(* IEC 61131-3 sources: CS_4_Aufzugsteuerung/src/Stations/CP112/Steuerung/Class/DiasMasterMain (part 2) *)

	l.eax		  RTCY
	and.eax		Dmrealtime
	call		  StoreNewPointers

END_FUNCTION
#endif

#ifdef _LSL_TARGETARCH_ARM
FUNCTION VIRTUAL GLOBAL DiasMasterMain::AddRet
  VAR_INPUT
    RTCY		: DINT;
  END_VAR

  if (RTCY AND DMREALTIME) = DMREALTIME then
    ud_DelayRealtime += C_TimeRet;
  else
    ud_DelayCyclic += C_TimeRet;
  end_if;

  (PtrCode + IPSub + RetStruct.Opc)^ := DbRet;

  IPSub += sizeof(RetStruct);

END_FUNCTION

#else
FUNCTION AWL VIRTUAL GLOBAL DiasMasterMain::AddRet
  VAR_INPUT
    RTCY		: DINT;
  END_VAR

	l.eax		  RTCY
	and.eax		Dmrealtime

//#SR001 Start
	CMP.EAX		Dmrealtime
	JNE			  LABEL_AR_NORT
	ADD.D		  ud_DelayRealtime,C_TimeRet
  JMP       LABEL_AR_TIMETAKEN

LABEL_AR_NORT
//#SR001 End
	ADD.D		  ud_DelayCyclic,C_TimeRet

LABEL_AR_TIMETAKEN

	call		  GetProgPointer

  l.ebx     PtrCode

	l.b			  (edx+ebx+RetStruct.Opc),DbRet			     // opcode Ret
	add.edx		sizeof (RetStruct)

	l.eax		  RTCY
	and.eax		Dmrealtime
	call		  StoreNewPointers

END_FUNCTION
#endif

//[English]
// Does a 16 Bit read access
//[Globals]		_RTOSVersion			: OS version
//				_lsl_pos				: OS interface structure
//[Members]
//[Locals]		ui_data			:R/W	:intermediate storeage of data
//				di_ret			:R/W	:returnvalue of OS
//[>Adress]		Module address and offset
//[<Data]		Data read
FUNCTION VIRTUAL GLOBAL DiasMasterMain::Rd16Bit
  VAR_INPUT
    Adress	: UDINT;
  END_VAR
  VAR_OUTPUT
    Data		: DINT;
  END_VAR
  VAR
    ui_data : uint;
    di_ret	: dint;
  END_VAR

	//ws005
	//*****************************************************
	//***** use OS functions instead of own functions *****
	//*****************************************************
	if( _RTOSVersion >= OSVersionDIASIO )then
		if( p_SemaHandle <> NIL )then			//ws007
			To_Multitask.Wait( p_SemaHandle );	//ws006
		end_if;
		di_ret := OS_DIAS_ReadWord( pDIAS  := pDIAS,
								   us_mod  := ( ( Adress shr 8 ) and 16#ff )$usint,
								   ui_off  := ( Adress and 16#ff )$uint,
								   ui_data := #ui_data );
		if( p_SemaHandle <> NIL )then				//ws007
			To_Multitask.Signal( p_SemaHandle );	//ws006
		end_if;
		if( di_ret <> 0 )then
			Data := 0;
			TraceAsyncError(( ( Adress shr 8 ) and 16#ff )$usint);
		else
			Data := ui_data;
		end_if;
	else
	//*****************************************************
	//*** use own functions (should be obsolete by now) ***
	//*****************************************************
	// /ws005
		TraceAsyncError(( ( Adress shr 8 ) and 16#ff )$usint);
	end_if;

END_FUNCTION

#ifdef _LSL_TARGETARCH_ARM
FUNCTION VIRTUAL GLOBAL DiasMasterMain::AddRd32Bit
  VAR_INPUT
    Adress		  : HINT;
    RTCY		    : DINT;
    thisp		    : ^void;
    callOptions : USINT;
  END_VAR
  VAR_OUTPUT
    Handle		  : DINT;
  END_VAR

  if (RTCY AND Dmrealtime) = Dmrealtime then
    ud_DelayRealtime += C_TimeRd8Bit + 3*(C_TimeRd16Bit - C_TimeRd8Bit); // appraised value: 1*basetime + 4*time for 1 byte (instead of C_TimeRd32Bit)
    ui_RtDIASAccesses += 1;
  else
    ud_DelayCyclic += C_TimeRd8Bit + 3*(C_TimeRd16Bit - C_TimeRd8Bit); // appraised value: 1*basetime + 4*time for 1 byte (instead of C_TimeRd32Bit)
    ui_CyDIASAccesses += 1;
  end_if;

  (PtrCode + IPSub + Rd32Struct.Opc)^         := DbRd32;
  (PtrCode$^HINT + IPSub + Rd32Struct.ChAdr)^ := Adress;

  ARM_EAX := RTCY$UDINT;
  ARM_EDI := thisp$UDINT;
  GetHandle(Rd32Struct.Data, callOptions);
  Handle := ARM_EAX$DINT;
  IPSub += sizeof(Rd32Struct);

END_FUNCTION

#else
// ***************************************
//   put programm into the buffer
// ***************************************
//  this is a 16 bit read
//  the thispointer we need to call the update method
//

FUNCTION AWL VIRTUAL GLOBAL DiasMasterMain::AddRd32Bit
	VAR_INPUT
		Adress 	    : HINT;
		RTCY 	      : DINT;
		thisp 	    : ^void;
		callOptions : USINT;
	END_VAR
	VAR_OUTPUT
		Handle 	    : DINT;
	END_VAR

	l.eax		  RTCY
	and.eax		Dmrealtime

//#SR001 Start
	CMP.EAX		Dmrealtime
	JNE			  LABEL_AR32B_NORT
	ADD.D		  ud_DelayRealtime,C_TimeRd32Bit
	inc.w		  ui_RtDIASAccesses
  JMP       LABEL_AR32B_TIMETAKEN

LABEL_AR32B_NORT
	ADD.D		  ud_DelayCyclic,C_TimeRd32Bit
	inc.w		  ui_CyDIASAccesses
//#SR001 End

LABEL_AR32B_TIMETAKEN

	call		  GetProgPointer

  l.ebx     PtrCode

	l.b			  (edx+ebx+Rd32Struct.Opc),DbRd32	   			// opcode Read 8
	l.ax		  Adress					// adress lo+high
	s.ax		  (edx+ebx+Rd32Struct.ChAdr+0)

	l.ax		  RTCY+0
	l.edi		  thisp				    // to put into then handle

  push.b    callOptions

	push.d		Rd16Struct.Data			// direct pointer on the data
	call		  GetHandle

  add.esp 5

	s.eax		  Handle

	add.edx		sizeof (Rd32Struct)

	l.eax		  RTCY
	and.eax		Dmrealtime
	call		  StoreNewPointers

END_FUNCTION
#endif

#ifdef _LSL_TARGETARCH_ARM
FUNCTION VIRTUAL GLOBAL DiasMasterMain::AddRd8Bit
  VAR_INPUT
    Adress		  : HINT;
    RTCY		    : DINT;
    thisp		    : ^void;
    callOptions : USINT;
  END_VAR
  VAR_OUTPUT
    Handle		  : DINT;
  END_VAR

  if (RTCY AND Dmrealtime) = Dmrealtime then
    ud_DelayRealtime += C_TimeRd8Bit;
    ui_RtDIASAccesses += 1;
  else
    ud_DelayCyclic += C_TimeRd8Bit;
    ui_CyDIASAccesses += 1;
  end_if;

  (PtrCode + IPSub + Rd8Struct.Opc)^         := DbRd8;
  (PtrCode$^HINT + IPSub + Rd8Struct.ChAdr)^ := Adress;

  ARM_EAX := RTCY$UDINT;
  ARM_EDI := thisp$UDINT;
  GetHandle(Rd8Struct.Data, callOptions);
  Handle := ARM_EAX$DINT;
  IPSub += sizeof(Rd8Struct);

END_FUNCTION

#else
// ***************************************
//   put programm into the buffer
// ***************************************
//  this is a 8 bit read
//  the thispointer we need to call the update method
//

FUNCTION AWL VIRTUAL GLOBAL DiasMasterMain::AddRd8Bit
	VAR_INPUT
		Adress 	    : HINT;
		RTCY 	      : DINT;
		thisp 	    : ^void;
		callOptions : USINT;
	END_VAR
	VAR_OUTPUT
		Handle 	    : DINT;
	END_VAR

	l.eax		  RTCY
	and.eax		Dmrealtime

//#SR001 Start
	CMP.EAX		Dmrealtime
	JNE			  LABEL_AR8B_NORT
	ADD.D		  ud_DelayRealtime,C_TimeRd8Bit
	inc.w		  ui_RtDIASAccesses			//#SR021
  JMP       LABEL_AR8B_TIMETAKEN

LABEL_AR8B_NORT
	ADD.D		  ud_DelayCyclic,C_TimeRd8Bit
	inc.w		  ui_CyDIASAccesses
//#SR001 End

LABEL_AR8B_TIMETAKEN

	call		  GetProgPointer

  l.ebx     PtrCode

	l.b			  (edx+ebx+Rd8Struct.Opc),DbRd8	   			// opcode Read 8
	l.ax		  Adress					// adress lo+high
	s.ax		  (edx+ebx+Rd8Struct.ChAdr+0)

	l.ax		  RTCY+0
	l.edi		  thisp				    // to put into then handle

  push.b    callOptions

	push.d		Rd8Struct.Data			// direct pointer on the data
	call		  GetHandle

  add.esp   5

	s.eax		  Handle
	add.edx		sizeof (Rd8Struct)

	l.eax		  RTCY
	and.eax		Dmrealtime
	call		  StoreNewPointers

END_FUNCTION
#endif

#ifdef _LSL_TARGETARCH_ARM
FUNCTION VIRTUAL GLOBAL DiasMasterMain::AddRTBSync
  VAR_INPUT
    Adress		: HINT;
  END_VAR
  VAR_OUTPUT
    FirstRTB	: DINT;
  END_VAR
  #ifdef OldDiasXilinx
  VAR
    pUSINT : ^USINT;
  END_VAR
#endif

  FirstRTB := 0;

  if DiasType <> 2 then

#IFNDEF OldDiasXilinx
    if RTBSyncAdr = NIL then
      RTBSyncAdr := (16#100*63+16#8002)$^USINT;// global sync

      FirstRTB := 1;
    end_if;
#ELSE
    if NumberSyncs >= NumberLocalSyncs then
      ErrorLocalSyncTrace();
    else
      ((#RtbLocalSyncAdr)$^DINT + NumberSyncs * (SIZEOF(RtbLocalSyncAdr)/NumberLocalSyncs))^ := Adress + 16#8000;
    end_if;
#ENDIF
  else
    // DiasType = 2 --> it is a new Master
#IFNDEF OldDiasXilinx
    if (SyncProgPtr + CntrlStruct.OPC)^ <> DbCntrl then
      (SyncProgPtr + CntrlStruct.OPC)^          := DbCntrl;
      (SyncProgPtr$^UINT + CntrlStruct.chAdr)^  := 16#100*63+2;
      (SyncProgPtr + CntrlStruct.Data)^         := 0;
      FirstRTB := 1;

      ud_DelayRealtime := ud_DelayRealtime + C_TimeControlWrite - C_TimeNop * 4; //because the 4 Nops were overwritten
    end_if;
#ELSE
    if NumberSyncs >= NumberLocalSyncs then
      ErrorLocalSyncTrace();
    else
      pUSINT := #CallsRt[0] + sizeof(TmrStruct) + NumberSyncs * SIZEOF(CntrlStruct);

      if (pUSINT + CntrlStruct.OPC)^ <> DbCntrl then
        (pUSINT + CntrlStruct.OPC)^         := DbCntrl;
        (pUSINT$^UINT + CntrlStruct.chAdr)^ := Adress;
        (pUSINT + CntrlStruct.Data)^        := 0;

        ud_DelayRealtime := ud_DelayRealtime + C_TimeControlWrite - C_TimeNop * 4; //because the 4 Nops were overwritten
      end_if;
    end_if;
#ENDIF
  end_if;

  NumberSyncs += 1;

  if FirstRTB = 1 then
    us_SyncModule := (Adress SHR 8)$USINT;
  end_if;

END_FUNCTION

#else

// *************************************************
//   RTB is fixed reserved for one MODUL
// *************************************************
//
//  if FirstRTB <> 0 then this modul is the first with RTB
//  and has to do perhaps something special
//  if FirstRTB = 0 then it already exists a modul with RTBSYNC
//

FUNCTION AWL VIRTUAL GLOBAL DiasMasterMain::AddRTBSync
  VAR_INPUT
    Adress		: HINT;
  END_VAR
  VAR_OUTPUT
    FirstRTB	: DINT;
  END_VAR

	l.d			FirstRTB,0

	cmp.b		DiasType,2			//ws005
	je			AddRTBIMaster		// --> it is a new Master

#IFNDEF OldDiasXilinx
	cmp.d		RTBSyncAdr,0
	jne			AddRTBSyncRet

	L.EDI		16#100*63+16#8002 		// global sync  //ws005: faster

	s.edi		RTBSyncAdr

	l.d			FirstRTB,1						// first RTB
#ELSE
	LZXW.EDI	Adress
	ADD.EDI		16#8000

	LZXB.EAX	NumberSyncs
	CMP.AL		NumberLocalSyncs
	JAE			  ErrorSync
	L.AH		  SIZEOF(RtbLocalSyncAdr)/NumberLocalSyncs
	MUL			  AH
	ADD.EAX		#RtbLocalSyncAdr

	S.EDI		  (EAX)
#ENDIF
	jmp			  AddRTBSyncRet

AddRTBIMaster
#IFNDEF OldDiasXilinx

	//#SR003 Start
	l.edi	    SyncProgPtr
	//#SR003 End

	cmp.b		  (edi+CntrlStruct.OPC),DbCntrl
	je			  AddRTBSyncRet

	l.b			  (edi+CntrlStruct.OPC),DbCntrl

	l.ax		  16#100*63+2 		// global sync

	s.ax		  (edi+CntrlStruct.chAdr+0)		// the modul normal = 63 (global SYNC)

	l.b			  (edi+CntrlStruct.Data),0		// we always write data 0
	l.d			  FirstRTB,1						// first RTB

//#SR001 Start
	SUB.D		  ud_DelayRealtime,C_TimeNop * 4			//because the 4 Nops were write over
	ADD.D		  ud_DelayRealtime,C_TimeControlWrite
//#SR001 End

#ELSE
	l.edi		  #CallsRt
	add.edi		sizeof (TmrStruct)  // the first INSTR is tmr

	LZXB.EAX	NumberSyncs
	CMP.AL		NumberLocalSyncs
	JAE			  ErrorSync
	L.AH		  SIZEOF(CntrlStruct)
	MUL			  AH
	ADD.EDI		EAX

	cmp.b		  (edi+CntrlStruct.OPC),DbCntrl
	je			  AddRTBSyncRet

	l.b			  (edi+CntrlStruct.OPC),DbCntrl
	l.ax		  Adress
	s.ax		  (edi+CntrlStruct.chAdr+0)		// the modul normal = 63 (global SYNC)

	l.b			  (edi+CntrlStruct.Data),0		// we always write data 0

//#SR001 Start
	SUB.D		  ud_DelayRealtime,C_TimeNop * 4			//because the 4 Nops were write over
	ADD.D		  ud_DelayRealtime,C_TimeControlWrite
//#SR001 End

	JMP			  AddRTBSyncRet

ErrorSync
	FC			  ErrorLocalSyncTrace
#ENDIF

AddRTBSyncRet

	INC.B		  NumberSyncs

	//#SR008 start
	cmp.d		  FirstRTB,1
	jne			  LABEL_End

	l.ax		  Adress
	shr.ax		8
	s.al		  us_SyncModule

LABEL_End
	//#SR008 end

END_FUNCTION
#endif

#ifdef _LSL_TARGETARCH_ARM
FUNCTION VIRTUAL GLOBAL DiasMasterMain::AddWR16Bit
  VAR_INPUT
    adress	    : Hint;
    RTCY		    : DINT;
    thisp		    : ^void;
    data		    : UINT;
    callOptions : USINT;
  END_VAR
  VAR_OUTPUT
    handle		  : DINT;
  END_VAR

  if (RTCY AND Dmrealtime) = Dmrealtime then
    ud_DelayRealtime += C_TimeWr16Bit;
    ui_RtDIASAccesses += 1;
  else
    ud_DelayCyclic += C_TimeWr16Bit;
    ui_CyDIASAccesses += 1;
  end_if;

  (PtrCode + IPSub + Wr16Struct.Opc)^         := DbWr16;
  (PtrCode$^HINT + IPSub + Wr16Struct.ChAdr)^ := Adress;
  (PtrCode$^HINT + IPSub + Wr16Struct.Data)^  := data;

  ARM_EAX := RTCY$UDINT;
  ARM_EDI := thisp$UDINT;
  GetHandle(Wr16Struct.Data, callOptions);
  Handle := ARM_EAX$DINT;
  IPSub += sizeof(Wr16Struct);

END_FUNCTION

// ***************************************
//   put programm into the buffer
// ***************************************
//  this is a 16 bit read
//  the thispointer we need to call the update method
//
#else
FUNCTION AWL VIRTUAL GLOBAL DiasMasterMain::AddWR16Bit
	VAR_INPUT
		adress 	      : HINT;
		RTCY 	        : DINT;
		thisp 	      : ^void;
		data 	        : UINT;
		callOptions 	: USINT;
	END_VAR
	VAR_OUTPUT
		handle 	      : DINT;
	END_VAR

	l.eax		  RTCY
	and.eax		Dmrealtime

//#SR001 Start
	CMP.EAX		Dmrealtime
	JNE			  LABEL_AW16B_NORT
	ADD.D		  ud_DelayRealtime,C_TimeWr16Bit
	inc.w		  ui_RtDIASAccesses			//#SR021
  JMP       LABEL_AW16B_TIMETAKEN

LABEL_AW16B_NORT
	ADD.D		  ud_DelayCyclic,C_TimeWr16Bit
	inc.w		  ui_CyDIASAccesses
//#SR001 End

LABEL_AW16B_TIMETAKEN

	call		  GetProgPointer

  l.ebx     PtrCode

	l.b			  (edx+ebx+Wr16Struct.Opc),DbWr16	   			// opcode Read 8
	l.ax		  Adress					// adress lo+high
	s.ax		  (edx+ebx+Wr16Struct.ChAdr+0)

	l.ax		  data
	s.ax		  (edx+ebx+Wr16Struct.Data)

	l.ax		  RTCY+0
	l.edi		  thisp				    // to put into then handle

  push.b    callOptions

	push.d		Wr16Struct.Data			// direct pointer on the data
	call		  GetHandle

  add.esp   5

	s.eax		  Handle

	add.edx		sizeof (Wr16Struct)
	l.eax		  RTCY
	and.eax		Dmrealtime
	call		  StoreNewPointers

END_FUNCTION
#endif

#ifdef _LSL_TARGETARCH_ARM
FUNCTION VIRTUAL GLOBAL DiasMasterMain::AddWr8Bit
	VAR_INPUT
		adress 	    : HINT;
		RTCY 	      : DINT;
		thisp 	    : ^void;
		Data 	      : USINT;
		callOptions : USINT;
	END_VAR
	VAR_OUTPUT
		Handle 	    : DINT;
	END_VAR

  if (RTCY AND Dmrealtime) = Dmrealtime then
    ud_DelayRealtime += C_TimeWr8Bit;
    ui_RtDIASAccesses += 1;
  else
    ud_DelayCyclic += C_TimeWr8Bit;
    ui_CyDIASAccesses += 1;
  end_if;

  (PtrCode + IPSub + Wr8Struct.Opc)^         := DbWr8;
  (PtrCode$^HINT + IPSub + Wr8Struct.ChAdr)^ := Adress;
  (PtrCode$^HINT + IPSub + Wr8Struct.Data)^  := data;

  ARM_EAX := RTCY$UDINT;
  ARM_EDI := thisp$UDINT;
  GetHandle(Wr8Struct.Data, callOptions);
  Handle := ARM_EAX$DINT;
  IPSub += sizeof(Wr8Struct);

END_FUNCTION

#else
FUNCTION AWL VIRTUAL GLOBAL DiasMasterMain::AddWr8Bit
	VAR_INPUT
		adress 	    : HINT;
		RTCY 	      : DINT;
		thisp 	    : ^void;
		Data 	      : USINT;
		callOptions : USINT;
	END_VAR
	VAR_OUTPUT
		Handle 	    : DINT;
	END_VAR

	l.eax		  RTCY
	and.eax		Dmrealtime

//#SR001 Start
	CMP.EAX		Dmrealtime
	JNE			  LABEL_AW8B_NORT
	ADD.D		  ud_DelayRealtime,C_TimeWr8Bit
	inc.w		  ui_RtDIASAccesses			//#SR021
  JMP       LABEL_AW8B_TIMETAKEN

LABEL_AW8B_NORT
	ADD.D		  ud_DelayCyclic,C_TimeWr8Bit
	inc.w		  ui_CyDIASAccesses
//#SR001 End

LABEL_AW8B_TIMETAKEN

	call		  GetProgPointer

  l.ebx     PtrCode

	l.b			  (edx+ebx+Wr8Struct.Opc),DbWr8	   			// opcode Read 8
	l.ax		  Adress					// adress lo+high
	s.ax		  (edx+ebx+Wr8Struct.ChAdr+0)
	l.al		  data
	s.al		  (edx+ebx+Wr8Struct.Data)

	l.ax		  RTCY+0
	l.edi		  thisp				    // to put into then handle

  push.b    callOptions

	push.d	  Wr8Struct.Data			// direct pointer on the data
	call		  GetHandle

  add.esp   5
	s.eax		  Handle

	add.edx		sizeof (Wr8Struct)

	l.eax		  RTCY
	and.eax		Dmrealtime
	call		  StoreNewPointers

END_FUNCTION
#endif

//[English]
// Function is writing into controlarea of a diasmodul
//[Globals]		_RTOSVersion		: OS version
//				_lsl_pos			: OS interface structure
//[Members]
//[Locals]
//[>Adress]		High Byte Modulnumber, Low Byte offset in Controlarea
//[>Data]		Data to write
//[<state]		0..success
FUNCTION VIRTUAL GLOBAL DiasMasterMain::WrCntr
  VAR_INPUT
    adress		: DINT;
    Data		  : Usint;
  END_VAR
  VAR_OUTPUT
    state		: DINT;
  END_VAR

	//ws005
	//*****************************************************
	//***** use OS functions instead of own functions *****
	//*****************************************************
	if( _RTOSVersion >= OSVersionDIASIO )then
		if( p_SemaHandle <> NIL )then			//ws007
			To_Multitask.Wait( p_SemaHandle );	//ws006
		end_if;
		state := OS_DIAS_WriteCtrl_( pDIAS  := pDIAS,
									us_mod  := ( ( Adress shr 8 ) and 16#ff )$usint,
									ui_off  := ( Adress and 16#ff )$uint,
									us_data := Data );
		if( p_SemaHandle <> NIL )then				//ws007
			To_Multitask.Signal( p_SemaHandle );	//ws006
		end_if;
		if( state <> 0 )then
			TraceAsyncError(( ( Adress shr 8 ) and 16#ff )$usint);
		end_if;
	else
	//*****************************************************
	//*** use own functions (should be obsolete by now) ***
	//*****************************************************
		if( ( _WhoAmI = 16#19 ) | ( _WhoAmI = 16#17 ) )then //ET261 and ETT321
			state := OS_DIAS_WriteCtrl_( pDIAS  := pDIAS,
										us_mod  := ( ( Adress shr 8 ) and 16#ff )$usint,
										ui_off  := ( Adress and 16#ff )$uint,
										us_data := Data );
			if( state <> 0 )then
				TraceAsyncError(( ( Adress shr 8 ) and 16#ff )$usint);
			end_if;
		else

	// /ws005
			TraceAsyncError(( ( Adress shr 8 ) and 16#ff )$usint);
		end_if;
	end_if;

END_FUNCTION
//[#ENGLISH]
//[>Time_uSec]Time in uSec (valid from 0-255)

#ifdef _LSL_TARGETARCH_ARM
FUNCTION VIRTUAL GLOBAL DiasMasterMain::AddWait
  VAR_INPUT
    RTCY		  : DINT;
    Time_uSec	: DINT;
  END_VAR

  if (RTCY AND Dmrealtime) = Dmrealtime then
    ud_DelayRealtime += Time_uSec$UDINT * 1000;
  else
    ud_DelayCyclic += Time_uSec$UDINT * 1000;
  end_if;

  (PtrCode + IPSub + DelayStruct.Opc)^       := DbDelay;
  (PtrCode + IPSub + DelayStruct.TIME_uSec)^ := Time_uSec$HSINT;

  IPSub += sizeof(DelayStruct);

END_FUNCTION
#else

FUNCTION AWL VIRTUAL GLOBAL DiasMasterMain::AddWait
  VAR_INPUT
    RTCY		  : DINT;
    Time_uSec	: DINT;
  END_VAR

	l.eax		  RTCY
	and.eax		Dmrealtime

//#SR001 Start
	l.ecx		  Time_usec
	imul.ecx	ecx,1000
	CMP.EAX		Dmrealtime
	JNE			  LABEL_AW_NORT
	ADD.D		  ud_DelayRealtime,ecx
  JMP       LABEL_AW_TIMETAKEN

LABEL_AW_NORT
  ADD.D		  ud_DelayCyclic,ecx
//#SR001 End

LABEL_AW_TIMETAKEN

	call		  GetProgPointer

  l.ebx     PtrCode

	l.b			  (edx+ebx+DelayStruct.OPC),DbDelay	   			// opcode delay uSec
	l.eax		  Time_uSec
	s.al		  (edx+ebx+DelayStruct.TIME_uSec)
	add.edx		sizeof (DelayStruct)

	l.eax		  RTCY
	and.eax		Dmrealtime
	call		  StoreNewPointers

END_FUNCTION
#endif

FUNCTION VIRTUAL GLOBAL DiasMasterMain::GetPllTime
  VAR_OUTPUT
    PllTime		: DINT;
  END_VAR
  VAR
    objinfo : LSLOBJ_INFO;
    Val		: DINT;
  END_VAR

	IF PllTimeGlob = 0 THEN

		To_TaskObjectControl.GetObjectInfo(this,OBJ_RT,#objinfo);			//#SR009

		// the set value of object
		PllTimeGlob := objinfo.period$DINT;
		IF PllTimeGlob = 0 THEN
#ifdef HWC_LogError
      HWC_LogError(this, "@0002 (DiasMasterMain::GetPllTime) A realtime of object 'DiasMasterC' is required !! ( 1ms is the default value ) !!");
#else
      TRACE("A realtime of object 'DiasMasterC' is required !! ( 1ms is the default value ) !!");
#endif
		END_IF;

    //look if we have µs or ms (µs msb is set)
    if ( ( objinfo.period and 16#8000_0000 ) = 0 ) then

      //we need our task time in µs
      ud_TaskTime := objinfo.period * 1000;
    else

      //we have already µs seconds
      ud_TaskTime := objinfo.period and 16#7FFF_FFFF;
    end_if;

		//#SR013 start
		us_RtPasses := 1;
		us_ModuleUpdate1ms := 1;
		us_MuSecMode := 0;

		//look if we have no old OS ( from 1.1.50 upwards)
		if _RtOSversion >= 16#1132 then
			//RTOS variable _ClockTicks ( with pointer because of linker error with old loaders without this variable)
			//_Firstscan has Offset 0EB8 and _ClockTicks has offset 0EAB, therefore -13
			ui_ClockTicks := ( ( #_Firstscan - 13 )$^UINT )^;

      if ui_ClockTicks < 1000 then
        //is DiasMaster rt time same as OS-Time (maintimer)
        if ( PllTimeGlob and 16#7FFF_FFFF ) = ui_ClockTicks then
          // check if maintimer has a valid value
          if ( 1000 mod ui_ClockTicks ) | ui_ClockTicks < 50 then
#ifdef HWC_LogError
            HWC_LogError(this, "@0003 (DiasMasterMain::GetPllTime) No valid maintimer value in OS (valid: 50,100,125,200,250,500,1000)! Master is set off!");
#else
            TRACE( "No valid maintimer value in OS (valid: 50,100,125,200,250,500,1000)! Master is set off!" );
#endif
            MasterOn := 0;
            ImOff := 1;
          else
            us_RtPasses := ( 1000 / ui_ClockTicks )$USINT;
            us_MuSecMode := 1;
            us_ModuleUpdate1ms := 0;
          end_if;
        else
          // there is only one FPGA SyncOut for OS-RT and DiasMaster, so they have to be at the same cycle
#ifdef HWC_LogError
          HWC_LogError(this, "@0004 (DiasMasterMain::GetPllTime) Rt-Time of DiasMasterC not the same as Base Rt-Time of OS (Maintimer). Master is set off!");
#else
          TRACE( "Rt-Time of DiasMasterC not the same as Base Rt-Time of OS (Maintimer). Master is set off!" );
#endif
          MasterOn := 0;
          ImOff := 1;
        end_if;
      end_if;
		end_if;
		//#SR013 End

		// but it could be a CPU with 3ms
		Val := PllTimeGlob MOD Ops.RtInterv_mSec$DINT;
		IF Val THEN
			PllTimeGlob += Ops.RtInterv_mSec$DINT - Val ;
		END_IF;

		// there could be a error
		IF PllTimeGlob < Ops.RtInterv_mSec$DINT THEN
			PllTimeGlob := Ops.RtInterv_mSec$DINT;
		END_IF;

#ifdef HWC_LogValue1
    HWC_LogValue1(this, "@0500 (DiasMasterMain::GetPllTime) PllTime = {0}", PllTimeGlob$UDINT);
#else
		//#SR008 start
		if p_KernelLog <> NIL then
			OS_KernelLog1( "DiasMaster: PllTime = %d", PllTimeGlob );
		end_if;
		//#SR008 end
#endif

		sd_PllTimeGlob_us := PllTimeGlob * 1000;		//#SR009
	END_IF;

	// aber eigentlich hängt er ja am TASK0 => #FA fragen !! => Ops.RtInterv_mSec

	PllTime := PllTimeGlob;

END_FUNCTION
//[English]
// Does a 8 Bit write access
//[Globals]		_RTOSVersion		: OS version
//				_lsl_pos			: OS interface structure
//[Members]
//[Locals]
//[>Adress]		Module address and offset
//[>Data]		Data to write
//[<State]
FUNCTION VIRTUAL GLOBAL DiasMasterMain::Wr8Bit
  VAR_INPUT
    Adress	: UDINT;
    Data		: Usint;
  END_VAR
  VAR_OUTPUT
    State		: DINT;
  END_VAR

	//ws005
	//*****************************************************
	//***** use OS functions instead of own functions *****
	//*****************************************************
	if( _RTOSVersion >= OSVersionDIASIO )then
		if( p_SemaHandle <> NIL )then			//ws007
			To_Multitask.Wait( p_SemaHandle );	//ws006
		end_if;
		State := OS_DIAS_WriteByte(pDIAS   := pDIAS,
                               us_mod  := ( ( Adress shr 8 ) and 16#ff )$usint,
                               ui_off  := ( Adress and 16#ff )$uint,
                               us_data := Data );
		if( p_SemaHandle <> NIL )then				//ws007
			To_Multitask.Signal( p_SemaHandle );	//ws006
		end_if;
		if( State <> 0 )then
			TraceAsyncError(( ( Adress shr 8 ) and 16#ff )$usint);
		end_if;
	else
	//*****************************************************
	//*** use own functions (should be obsolete by now) ***
	//*****************************************************
	// /ws005
		TraceAsyncError(( ( Adress shr 8 ) and 16#ff )$usint);
	end_if;

END_FUNCTION

FUNCTION  DiasMasterMain::DiasMasterMain
  VAR_OUTPUT
    ret_code		: CONFSTATES;
  END_VAR
  VAR
    MyProgPtr       : ^USINT;
    P2Cil		        : ^s_DiasInfoType;	//ws003
    i		            : USINT;
    PTRWDDIAS	      : ^USINT;
    SigmaTekDevInfo : ^PCICONFDATA;
    timex		        : UDINT;
#ifndef HWC_LogInit
    P2SSR		        : ^LSL_SSR;				//#SR008
#endif
    p_Obj           : ^Obj;
    p_ClsHdr        : ^ClsHdr;
    b_IsLocalMaster : BOOL;
  END_VAR

  // check if we are any kind of derivation that makes us no local master!
  b_IsLocalMaster := TRUE;
  p_Obj		:= LSL_GetHdr(this);
  p_ClsHdr := p_Obj^.pClsHdr;
  WHILE p_clsHdr^.pBaseCls <> NIL DO // go down until there is no base - we might be derived by the user....
    #pragma warning(disable: 137 )
    IF  _strcmp(str1:=#p_ClsHdr^.pDsc^.Name.Text$CHAR, str2:="Dias2DataMover") = 0
      | _strcmp(str1:=#p_ClsHdr^.pDsc^.Name.Text$CHAR, str2:="DiasMasterSplitter") = 0
      | _strcmp(str1:=#p_ClsHdr^.pDsc^.Name.Text$CHAR, str2:="DiasMasterC_Dummy") = 0 THEN
      //if we find a derivation during going down that is called Dias2DataMover or DiasMasterSplitter
      //this is no local DiasMaster and we do not need to initialize it
      b_IsLocalMaster := FALSE;
      EXIT;
    END_IF;
    #pragma warning(default: 137 )
    p_ClsHdr := p_ClsHdr^.pBaseCls;
  END_WHILE;

  MasterON := 1;
  RTBSyncAdr :=NIL;
  CDiasType:=0;
  DiasType := 16#ff;
  ud_DelayRealtime := 0;	//#SR001
  us_SyncModule := 255;	//#SR012

  //#SR013 start
  us_RtPasses := 1;
  us_ModuleUpdate1ms := 1;
  us_MuSecMode := 0;
  //#SR013 end

  PtrCY 	 := #CallsCY[0];
  IPMainCY := 0;   // stops with a end programm
  IPSub  := 0;//(DmCallRes* sizeof (CallStruct)) + sizeof (EndStruct);

  PtrRT 	 := #CallsRT[0];

  PtrCode  := #CodeRtCy[0];

  IF b_IsLocalMaster THEN

    pDIAS := _lsl_pos^.piDias;  //ws005: prepare the DIAS pointer (faster)

#ifdef HWC_LogInit
    HWC_LogInit();
#else
    //#SR008 start
    if OS_CILGET( "SSR", #P2SSR ) then
      p_KernelLog := NIL;
    else
      p_KernelLog := ( P2SSR^.KernelLog )$^DINT;
    end_if;
    //#SR008
#endif

    // test if interface already exist
    if OS_CILGET("DiasInfo", #P2Cil) then
      if ((_IOsegment$DINT <> 0) & (_IOsegment$DINT <> 16#D0000)) then
        release :=0;
        DiasType:=1;
      end_if;
    else
      DiasType := P2Cil^.DiasType$usint;
      _IOSegment$^USINT := DiasHwPointer  := P2Cil^.DiasHWPointer$^usint; //ws003
      CDiasHwPointer := P2Cil^.CDiasHWPointer$^usint;	//ws003
      CDiasType := ( P2Cil^.CDiasType )$USINT;	//ws003

      IF CDiasType = 1 THEN

        //--- CCL -----------------------------------------------------
        IF OS_CILGET("CDIAS_IRQ",#lsl_cdias_irq) = SYS_ERR_NONE THEN
          CDiasIRQpossible := 1;
        END_IF;

      ELSIF CDiasType = 2 THEN

        //--- CIPC ----------------------------------------------------
        IF OS_CILGET("CDIAS_IRQ",#lsl_cdias_irq) = SYS_ERR_NONE THEN
          CDiasIRQpossible := 1;
        END_IF;

        IF OS_CILGET("PCICONFIG", #pSPCIInfo) =  SYS_ERR_NONE THEN
          // watchdog C-DIAS Bus
          // Trigger: write on offset 13 value 0
          SigmaTekDevInfo := SPCIINFO_FINDDEVICEBYNAME( "CDIASWATCHDOG" ,0 );
          CDiasI2CWatchdog$pVoid := SPCIINFO_GETADDRESS(SigmaTekDevInfo);
          CDiasI2CWatchdog$UDINT += 13;
          CDiasI2CWatchdog^ := 0;
          // #BS000
          i := (CDiasI2CWatchdog+2)^; // quit overrun (for Watchdog tracemessage)
        ELSE
#ifdef HWC_LogError
          HWC_LogError(this, "@0005 (DiasMasterMain::DiasMasterMain) A newer OS is required to insure a correct functionality of the CDIAS-Bus of the CPU !!");
#else
          Trace("A newer OS is required to insure a correct functionality of the CDIAS-Bus of the CPU !!");
#endif
        END_IF;

        //#SR016 start
        if ( P2Cil^.PLLType = 2 ) then

          //get pointer to new pll
          p_NewPll$^UDINT := ( P2Cil^.PLLHWPointer )$^UDINT;
        else
        //#SR016 end

          // sync on cdias bus
          CDIASSync$UDINT := P2Cil^.PLLHWPointer;		//ws003
          (CDIASSync+1)^ := ops.RtInterv_mSec$USINT; // Set Sync Time on CDIAS-Bus
        end_if;			//#SR016

      END_IF;
    end_if;

    // on linux platforms there is no local DIAS/CDIAS
    if ops_is_linux() = 0 then
      if _WHOAMI <= 16#35 then  //LanSte 09.12.2013 Only check for relativly old CPU's, newer CPU's may have no DIAS Bus at all.
        if (DiasType = 16#2) | (DiasType = 16#ff) then
          if TestMasterIM() = TRUE then
            // #BS 240903
            PTRWDDIAS$UDINT := _IOSegment$UDINT + DMWDTriggerMode;
            PTRWDDIAS^ := 0; // set to Trigger on async too
            PTRWDDIAS$UDINT := _IOSegment$UDINT + DMWDTimeBase;
            PTRWDDIAS^ := 8; // set timebase of watchdog to 8*16=128ms

            DiasType:=2;		// we are a IMaster
            InitChip();

            // to skip DiasError 63 on old intellgent master
            // #BS007
            timex := ops.tAbsolute;
            WHILE ops.tAbsolute - timex <= 150ms DO END_WHILE;
          else
              // if IOsegment <> 0 then it must be a old standard master
            if _IOsegment <> 0 then
              release :=0;
              DiasType:=1;
            end_if;

          END_IF;
        end_if;
      else
        Release   := 16#FFFFFFFF;   // Fehler Master nicht vorhanden
        MasterON  := 0;
      end_if;
    else
      Release   := 16#FFFFFFFF;   // Fehler Master nicht vorhanden
      MasterON  := 0;
    end_if;
  // pointer to top of programm and we keep space for 100 calls + END

  // 1. in the RT Prog at the begin is fix wait timer event

    #IFNDEF OldDiasXilinx

    //#SR013 start
    IPMainRT := sizeof( EventStruct );
  #ELSE
    i := NumberLocalSyncs;
    IF i THEN
      IPMainRT := sizeof (CntrlStruct) * NumberLocalSyncs + sizeof (EventStruct);
    ELSE
      IPMainRT := sizeof (CntrlStruct) + sizeof (EventStruct);
    END_IF;

  #ifdef HWK_SHOW_PRAGMA_MESSAGES
      #pragma message("Hier wurde Code temporär von FucHer am 05.06.2013 16:38 geändert! Zurückbauen nicht vergessen!")
  #endif
  #ENDIF

    // always begins with a timer event and fixed NOP for SYNC

    MyProgPtr :=PtrRT;

    #pragma warning( disable: 74 )				//#SR007
    // timer event
    MyProgPtr^   := DbTmrEve;     // always at the begin is a timer event
    MyProgPtr    += 1;
    #pragma warning( default: 74 )				//#SR007

    ud_DelayRealtime += C_TimeTimerEvent;		//#SR001

    #IFNDEF OldDiasXilinx
    // control write = 4 Byte filled with nop's
    // only one global sync

    //#SR013 start
    if DiasType =  2 then
      AddCall2Main( Mode := DmSingle, RTCY := DMRealtime, thisp := NIL ); 	// pointer is set later
      SyncProgPtr$UDINT := IPSub$UDINT + ( #CodeRtCy )$UDINT;
      AddNOP( RTCY := DMRealtime, nCount := 4 );
      AddRet( RTCY := DMRealtime );

      HandleNrRt := 1;
    else
      HandleNrRt := 0;
    end_if;

    IPMainRT += 2 * sizeof( MoveStruct );
    MyProgPtr += sizeof( CallStruct );
    //#SR013

    //#SR010 start
    //Mark realtime task of intelligent master as active to find out if realtime is already running when
    //Rt of DiasMasterC starts (Byte is only read in DiasMasterC Rt - Program)
    MyProgPtr^	:= DbMov;
    MyProgPtr   += 1;
    ( MyProgPtr$^UINT )^	:= DmUserData + 1;
    MyProgPtr   += 2;
    ( MyProgPtr$^UINT )^	:= DmUserData + 3;
    MyProgPtr	+= 2;

    ud_DelayRealtime += C_TimeMove;

    //Set Bit to recognize that realtime of IM doesn't start when Rt of DiasMaster runs
    //(Byte is reseted at the beginning of DiasMasterC Rt - Program)
    MyProgPtr^	:= DbMov;
    MyProgPtr	+= 1;
    ( MyProgPtr$^UINT )^	:= DmUserData + 1;
    MyProgPtr	+= 2;
    ( MyProgPtr$^UINT )^	:= DmUserData + 4;

    ud_DelayRealtime += C_TimeMove;

    //save copy values in UserData Area
    if( DiasType = 2 )then
      MyProgPtr 	:= ( _IOSegment + DmUserData + 1 )$^USINT;
      MyProgPtr^	:= 1;
      MyProgPtr	+= 1;
      MyProgPtr^	:= 0;
    end_if;
    //#SR010 end

  #ELSE
    // many local syncs
    i := NumberLocalSyncs;
    IF i THEN
      FOR i := 0 TO NumberLocalSyncs-1 DO
        MyProgPtr^   := DbNOP;
        MyProgPtr    += 1;
        MyProgPtr^   := DbNOP;
        MyProgPtr    += 1;
        MyProgPtr^   := DbNOP;
        MyProgPtr    += 1;
        MyProgPtr^   := DbNOP;
        MyProgPtr    += 1;
      END_FOR;

      ud_DelayRealtime += ( C_TimeNop	* 4 * NumberLocalSyncs );	//#SR001

    ELSE
      // we say 1 sync is required
      MyProgPtr^   := DbNOP;
      MyProgPtr    += 1;
      MyProgPtr^   := DbNOP;
      MyProgPtr    += 1;
      MyProgPtr^   := DbNOP;
      MyProgPtr    += 1;
      MyProgPtr^   := DbNOP;
      MyProgPtr    += 1;

      ud_DelayRealtime += ( C_TimeNop	* 4 );	//#SR001

    END_IF;
    HandleNrRt := 0;		//#SR013
  #ENDIF

    //get interface for hardwaretree functions
    if ( OS_CILGET(INTERFACE_HARDWARETREE, #pHardwareTree)) then
      pHardwareTree := NIL;

#ifdef HWC_LogError
      HWC_LogError(this, "@0006 (DiasMasterMain::DiasMasterMain) Hardwaretree-Interface not found. A newer OS is required for Safety-Modules");
#else
      TRACE("Hardwaretree-Interface not found. A newer OS is required for Safety-Modules");
      if p_KernelLog <> NIL then
        OS_KernelLog0("Hardwaretree-Interface not found. A newer OS is required for Safety-Modules");
      end_if;
#endif
    end_if;

    HandleNrCy := 0;

    ReadAllKenn();  // must be done in the constructor

  END_IF;

  ret_code	:= C_OK;

END_FUNCTION

#ifdef _LSL_TARGETARCH_ARM
FUNCTION DiasMasterMain::InitChip
  VAR
    Temp : DINT;
  END_VAR

// *****************************************
//  all programms off and chip on risk off
// *****************************************

  (_IOSegment$^USINT + DmControl)^  :=  1;  // Chip On, Risc Off
  (_IOSegment$^USINT + DmState)^    :=  0;  // All Programms OFF

// **********************************************
//  set period time of PLL
// **********************************************

// Pll Periode is overwritten later by realtime time of object
  (_IOSegment$^USINT + DmPllSyncDel)^  :=  (1000/DmTmrResso - 975/DmTmrResso);
  (_IOSegment$^USINT + DmPllPeriode)^  :=  ops.RtInterv_mSec$USINT;

// ****************************************************
//  we divide the complete memory into 3 fixed parts (1/4 for Cy Calls, 1/4 for Rt Calls and 1/2 for RtCy Code)
// ****************************************************

  (_IOSegment$^UINT + DmCyStartAdrM0)^   := 0; // Cyclic Start at Adr 00

  ud_IMMemory := (((_IOSegment$^USINT + DmCR_ProgMem)^ SHR 1) SHL 10);  // wieviel programm speicher haben wir
  (_IOSegment$^UINT + DmRtStartAdrM0)^ := (ud_IMMemory SHR 2)$UINT;

// *********************************
//  mov the IP to start destination
// *********************************

  StartOfCode := ud_IMMemory$DINT SHR 1;  // we use 2nd half of memory for the code => divide memory by 2

  Temp := (_IOSegment$^UINT + DmCyStartAdrM0)^;
  (_IOSegment$^UINT + DmCyProgCntrM0)^ := Temp$UINT; // CycPrgCntr = CycStart
  StartOfCy := Temp;

  Temp := (_IOSegment$^UINT + DmRtStartAdrM0)^;
  (_IOSegment$^UINT + DmRtProgCntrM0)^ := Temp$UINT; // RtPrgCntr = RtStart
  StartOfRt := Temp;

  (_IOSegment$^USINT + DmControl)^     := 2#11;   // Chip On, Risc On

END_FUNCTION
#else
FUNCTION  AWL DiasMasterMain::InitChip

  L.EDI      _IOSegment

// *****************************************
//  all programms off and chip on risk off
// *****************************************

	L.B		    (EDI+DmControl),1		// Chip On, Risc Off
	L.B		    (EDI+DmState)  ,0	    // All Programms OFF

// **********************************************
//  set period time of PLL
// **********************************************

	L.B		    (EDI+DmPllSyncDel),(1000/DmTmrResso  - 975/DmTmrResso)

// is overwritten later by realtime time of object
	L		      Ops.RtInterv_mSec+0		// Set Pll Periode
	S		      (EDI+DmPllPeriode)

// ****************************************************
//  we divide the complete memory into 3 fixed parts (1/4 for Cy Calls, 1/4 for Rt Calls and 1/2 for RtCy Code)
// ****************************************************

	L.W			  (EDI+DmCyStartAdrM0), 0   // Cyclic Start at Adr 00

	LZXB.eAX	(EDI+DmCR_ProgMem)		// wieviel programm speicher haben wir
	shr.eax		1									//#SR004
  shl.eax		8
	s.ax		  (EDI+DmRtStartAdrM0)
  shl.eax		2									//#SR004
	s.eax		  ud_IMMemory							//#SR004

// *********************************
//  mov the IP to start destination
// *********************************

  shr.eax   1  // we use 2nd half of memory for the code => divide memory by 2
  s.eax     StartOfCode

	LZXW.EAX	(EDI+DmCyStartAdrM0)
	S.AX		  (EDI+DmCyProgCntrM0)     // CycPrgCntr = CycStart
	s.eax		  StartOfCy

	LZXW.EAX	(EDI+DmRtStartAdrM0)
	S.AX		  (EDI+DmRtProgCntrM0)     // RtPrgCntr = RtStart
	s.eax		  StartOfRt

	L.B			  (EDI+DmControl),3	   // Chip On, Risc On

END_FUNCTION
#endif

//[English]
// reads all identification codes
//[Globals]		_RTOSVersion		:R		:OS version
//				_DiasConfig			:R/W	:configuration array (filled by OS)
//				_WhoAmI				:R		:CPU identification
//				OPS					:R		:OS variable
//[Members]		FirstModuleFound	:W		:determine a place on the bus where a modules is connected
//			(s) Release				:R		:Hardware + Software release
//[Locals]		MyTAbsolute			:R/W	:for a fixed time delay
FUNCTION  DiasMasterMain::ReadAllKenn
  VAR
    i           : usint;		//ws005
    MyTabsolute : DINT;
  END_VAR

	//ws005
	//*****************************************************
	//***** use OS functions instead of own functions *****
	//*****************************************************
	if( _RTOSVersion >= OSVersionDIASIO )then
		FirstModulFound := 16#ff;				//ws005
		for i := 0 to 62 do
			if( _DiasConfig[ i ] <> 255 )then 	// read directly from the DiasConfig
				FirstModulFound := i;           // which is provided by the OS
			end_if;								// this is in fact the last module in the array => does not matter
		end_for;
	else
	//*****************************************************
	//*** use own functions (should be obsolete by now) ***
	//*****************************************************
	// /ws005
		if Release <> 16#ffffffff then
			//ws004
			if( ( _WhoAmI = 16#19 ) | ( _WhoAmI = 16#17 ) )then //ET261 and ETT321

				FirstModulFound := 16#ff;	//ws005
				for i := 0 to 62 do
					if( _DiasConfig[ i ] <> 255 )then 	// read directly from the DiasConfig
						FirstModulFound := i;           // which is provided by the OS
					end_if;								// this is in fact the last module in the array => does not matter
				end_for;

			else
			// /ws004
				// dummy weil bus noch nicht laufen könnte
				ReadKenn(0);
				MyTabsolute := OPS.tAbsolute$DINT;
				while ((OPS.tabsolute - MyTabsolute$udint) < 50) do	//ws008
				end_while;;
				ReadKenn(0);

				// ************************************************
				// jetzt laufen alle Karten sicher
				// und darum können wir jetzt die Kennung lesen
				// ************************************************

				FirstModulFound := 16#ff;	//ws005

				For i:=0 to 62 do
					_Diasconfig[i] := to_USINT(ReadKenn(i));
					if _Diasconfig[i] <> 255 then
						FirstModulFound :=i;
					end_if;
				end_for;

				_Diasconfig[63]:=16#FF;  // sicher nicht da
				Return;

			end_if;

		else
		// otherwise you get problem on old DiasMasterMain + disable master = offline
			FirstModulFound :=16#FF;
			For i:=0 to 62 do
				_Diasconfig[i] := 16#FF;
			end_for;
		end_if;
	end_if;

END_FUNCTION
//[English]
// reads the identification code of one module
//[Globals]		_RTOSVersion		:R		:OS version
//				_lsl_pos			:R		:OS interface structure
//[Members]
//[Locals]
//[>Place]		Place on bus
//[<Kenn]		ID code
#pragma warning (disable:73)
#pragma warning (disable:76)
FUNCTION DiasMasterMain::ReadKenn
  VAR_INPUT
    Place		: DINT;
  END_VAR
  VAR_OUTPUT
    Kenn		: DINT;
  END_VAR
#ifdef _LSL_TARGETARCH_X86

	if( ImOff = 1 )then // Master is off
		Kenn := 16#ff;
		return;
  	end_if;

	//ws005
	//*****************************************************
	//***** use OS functions instead of own functions *****
	//*****************************************************
	if( _RTOSVersion >= OSVersionDIASIO )then
		if( pDIAS = NIL )then // OS has no Dias Interface (for now only CCL081)
			Kenn := 16#ff;
			return;
		end_if;
		Kenn := OS_DIAS_ReadKenn( pDIAS, Place$usint ); // OS function suits best
	else
	//*****************************************************
	//*** use own functions (should be obsolete by now) ***
	//*****************************************************
	// /ws005
		if( ( _WhoAmI = 16#19 ) | ( _WhoAmI = 16#17 ) )then //ET261 and ETT221
			Kenn := OS_DIAS_ReadKenn( pDias, Place$usint ); // OS function suits best
		else	//compatible mode
			TraceAsyncError(Place$usint);
		end_if;
  end_if;
#endif

END_FUNCTION
#pragma warning (default:73)
#pragma warning (default:76)
// /ws004

//[#ENGLISH]
//Diese Funktion prüft ob der Master vorhanden ist und wenn ja trägt Sie
//die HW und Software Kennung in Release ein
//
//IPC: (Hardware and software release)
//Bit 0-15   in Release ist Software Version // #BS016
//Bit 16-31  in Release ist Hardware Version
//
//C-IPC: (only one vlaue for hardware and software release)
//Bit 0-7
//
//Release = 16#FFFFFFFF ( Fehler Master nicht vorhanden)
//
//
#ifdef _LSL_TARGETARCH_ARM
FUNCTION DiasMasterMain::TestMasterIM
  VAR_OUTPUT
    MasterOK		: UINT;
  END_VAR

#ifndef DIAS_MASTER_PCI

  MasterOK := FALSE;
  Release := 16#FFFFFFFF;

  if DiasType <> 2 then                     // --> bereits erkannt über schnittstelle
    //---- Das Macht Später das BetrSyst !!---
    To_OSKernel.OutWord(Portnumber:=16#210, value:=(_IOSegment SHR 4)$UINT);  // Den CHIP In Den I/O Bereich legen
    To_OSKernel.OutByte(Portnumber:=16#212, value:=1);                        // Turn Chip
    if To_OSKernel.InWord(Portnumber:=16#21E) <> 16#494D then                 // "IM"
      return;
    end_if;
  end_if;

#endif

  if (_IOSegment$^UINT + DMID)^ <> 16#494d then // "IM"
    return;
  end_if;

  if CDiasType = 2 then
    Release := GetVerIMCIPC();
  else
    Release := (_IOSegment$^USINT + DMXVER)^;
  end_if;

  (_IOSegment$^USINT + DMCMDBUF1)^ := 3;  // Command Buffer Init mit Error
  (_IOSegment$^USINT + DMCMDBUF2)^ := 3;  // Command Buffer Init mit Error
  MasterOK := TRUE;

END_FUNCTION
#else
FUNCTION AWL  DiasMasterMain::TestMasterIM
  VAR_OUTPUT
    MasterOK		: UINT;
  END_VAR

#ifdef DIAS_MASTER_PCI
//
//	THR Aug. 21, 2003
//	To get a plug-in PCI card to work at D0000, bypass the "port"
//	test!!!
//	only on PC's with PCI412 and PCI402

	jmp				TestMasterGo
//
#endif	// DIAS_MASTER_PCI

	l.w			  MasterOK,FALSE
	l.d			  Release,16#ffffffff  	// Error

	cmp.b		  DiasType,2				//ws005
	je			  TestMasterGo			// --> bereits erkannt über schnittstelle

//---- Das Macht Später das BetrSyst !!---

	L.DX		  16#210					// Den CHIP In Den I/O Bereich Legen
	L.EAX		  _IOSegment
	SHR.EAX		4
	OUTW

	L.DX		  16#212					// Turn Chip
	L			    16#01
	OUTB

	l.dx		  16#21E
	inw
	cmp.ax 		16#494d					// "IM"
	jne			  TestMasterIMError		// --> no intelligent Master

//----------------------

TestMasterGo
	l.EDI		  _IOSegment
	l.ax 		  (EDI+DmID)
	cmp.ax 		16#494d					// "IM"
	jne			  TestMasterIMError
	CMP.b		  CDiasType,2 // #BS 100903	//ws005
	JE			  CIPCRelease

	// 	IPC
	clr			  eax
	l			    (EDI+DmXver)			// Xilinx  Version
	JMP			  CMDInitError

CIPCRelease
// #BS 100903 for C-IPC
	FC			  GetVerIMCIPC

CMDInitError
	s.eax		  Release

	l.b			  (EDI+DmCmdBuf1),3			// Command Buffer Init mit Error		//#SR017
	l.b			  (EDI+DmCmdBuf2),3			// Command Buffer Init mit Error 		//#SR017
	l.w			  MasterOK,TRUE

TestMasterIMError

END_FUNCTION
#endif
//
// --> ebx is this pointer
//     edx is IPSUB
//     ecx is IPMAIN
// --> ax mode reg  bit 0  = RT or Cyclic
//        			bit 14 =
// 					bit 15 = Main or Sub
//     edi thispointer
//
// <-- EAX is handle it is a direct pointer to the programm in the master
//

#ifdef _LSL_TARGETARCH_ARM
FUNCTION DiasMasterMain::GetHandle
  VAR_INPUT
    Offset        : UDINT;
    callOptions 	: USINT;
  END_VAR
  VAR
    pHandle       : ^OneHandle;
    SizeRtPostScan: DINT;
    SizeRt        : DINT;
    SizeCy        : DINT;
  END_VAR

  if ARM_EAX AND DmRealtime then
    // ** we put it into the realtime handlers **
    if callOptions AND CALL_OPTION_RT_POSTSCAN then
      SizeRtPostScan := HandleNrRtPostScan * sizeof(OneHandle);

      if SizeRtPostScan >= sizeof(HandlesRTPostScan) then
        //BLEERN - let the system crash if we try to allocate too many handles!
        pHandle$UDINT :=  0;
        pHandle$^UDINT^ := 0;
      end_if;

      pHandle := #HandlesRTPostScan[0] + SizeRtPostScan;
      pHandle^.Typ   := ARM_EAX$UINT;
      pHandle^.thisp := ARM_EDI$^HwBase;

      if ARM_EAX AND DmCallProg then    // test if it is Main Prog
        pHandle^.Address := (IPMainRT + StartOfRt + Offset$DINT)$UINT;
        ARM_EAX := pHandle^.Address;
      else
        pHandle^.Address := (IPSub + StartOfCode + Offset$DINT)$UINT;
        ARM_EAX := pHandle^.Address;
      end_if;

      HandleNrRtPostScan += 1;
    end_if;

    if callOptions AND CALL_OPTION_RT_PRESCAN then
      SizeRt := HandleNrRt * sizeof(OneHandle);

      if SizeRt >= sizeof(HandlesRT) then
        //BLEERN - let the system crash if we try to allocate too many handles!
        pHandle$UDINT :=  0;
        pHandle$^UDINT^ := 0;
      end_if;

      pHandle := #HandlesRT[0] + SizeRt;
      pHandle^.Typ   := ARM_EAX$UINT;
      pHandle^.thisp := ARM_EDI$^HwBase;

      if ARM_EAX AND DmCallProg then  // test if it is Main Prog
        pHandle^.Address := (IPMainRT + StartOfRt + Offset$DINT)$UINT;
        ARM_EAX := pHandle^.Address;
      else
        pHandle^.Address := (IPSub + StartOfCode + Offset$DINT)$UINT;
        ARM_EAX := pHandle^.Address;
      end_if;

      HandleNrRT += 1;
    end_if;

  else
    // ** we put it into the Cyclic handlers **
    SizeCy := HandleNrCY * sizeof(OneHandle);

    if SizeCy >= sizeof(HandlesCY) then
      //BLEERN - let the system crash if we try to allocate too many handles!
      pHandle$UDINT :=  0;
      pHandle$^UDINT^ := 0;
    end_if;

    pHandle := #HandlesCY[0] + SizeCy;
    pHandle^.Typ   := ARM_EAX$UINT;
    pHandle^.thisp := ARM_EDI$^HwBase;

    if ARM_EAX AND DmCallProg then  // test if it is Main Prog
      pHandle^.Address := (IPMainCY + StartOfCy + Offset$DINT)$UINT;
      ARM_EAX := pHandle^.Address;
    else
      pHandle^.Address := (IPSub + StartOfCode + Offset$DINT)$UINT;
      ARM_EAX := pHandle^.Address;
    end_if;

    HandleNrCY += 1;
  end_if;

END_FUNCTION
#else
FUNCTION AWL DiasMasterMain::GetHandle
	VAR_INPUT
		Offset 	    : UDINT;
		callOptions : USINT;
	END_VAR
  VAR
  	mode        : UDINT;
    old_ecx     : UDINT;
  END_VAR

	push		  edx
	push		  ecx

	clr			  ebx

  s.ecx     old_ecx

  s.eax     mode

	test.ax		Dmrealtime						// test if it is a realtime handle or not
	jnz			  GetHandleRTPostScan						// --> it is a realtime handle

// ** we put it into the Cyclic handlers **

	lzxw.ebx	HandleNrCY

//BLEERN - let the system crash if we try to allocate too many handles!
  cmp.ebx   (SIZEOF(HandlesCY) / SIZEOF(OneHandle))
  jne       HandleCyOK
  xor.edi   edi
  l.w       (edi), 0
HandleCyOK
//END BLEERN - let the system crash if we try to allocate too many handles!

  imul.ebx	ebx, sizeof (OneHandle)
	push		  edi
	l.edi		  #handlescy					   // there is an compiler error
	add.ebx	  edi							   // this is the reason wy we do this different
	pop			  edi

	s.ax		  (ebx+OneHandle.Typ)
	s.edi		  (ebx+OneHandle.thisp)

	test.ax		DmCallProg	    				// test if it is Main Prog
	jz			  getHandleCySB
	add.ecx		StartOfCy
	add.ecx		offset
	s.cx		  (ebx+OneHandle.Address)
	l.eax		  ecx
	jmp			  getHandleCyMain

getHandleCySB
	add.edx		StartOfCode
	add.edx		offset
	s.dx		  (ebx+OneHandle.Address)
	l.eax		  edx
getHandleCyMain

	inc.w		  HandleNrCY

	jmp			  GetHandleRet

// ** we put it into the realtime handlers **

GetHandleRTPostScan

  test.     b callOptions, CALL_OPTION_RT_POSTSCAN
  jz        GetHandleRT

  lzxw.ebx	HandleNrRtPostScan

//BLEERN - let the system crash if we try to allocate too many handles!
  cmp.ebx   (SIZEOF(HandlesRTPostScan) / SIZEOF(OneHandle))
  jne       HandleRTPostScanOk
  xor.edi   edi
  l.w       (edi), 0
HandleRTPostScanOK
//END BLEERN - let the system crash if we try to allocate too many handles!

	imul.ebx	ebx, sizeof (OneHandle)
	push		  edi
	l.edi		  #HandlesRTPostScan					   // there is an compiler error
	add.ebx		edi							   // this is the reason wy we do this different
	pop			  edi

	s.ax		  (ebx+OneHandle.Typ)
	s.edi		  (ebx+OneHandle.thisp)

	test.ax		DmCallProg						// test if it is Main Prog
	jz			  getHandleRtPostScanSB
	add.ecx		StartOfRt
	add.ecx		offset
	s.cx		  (ebx+OneHandle.Address)
	l.eax		  ecx								// handle
	jmp			  getHandleRtPostScanMain

getHandleRTPostScanSB
	add.edx		StartOfCode
	add.edx		offset
	s.dx		  (ebx+OneHandle.Address)
	l.eax		  edx

getHandleRtPostScanMain
	inc.w		  HandleNrRTPostScan

GetHandleRT

  test.b    callOptions, CALL_OPTION_RT_PRESCAN
  jz        GetHandleRet

  l.eax     mode
  l.ecx     old_ecx

  lzxw.ebx	HandleNrRt

//BLEERN - let the system crash if we try to allocate too many handles!
  cmp.ebx   (SIZEOF(HandlesRT) / SIZEOF(OneHandle))
  jne       HandleRTOk
  xor.edi   edi
  l.w       (edi), 0
HandleRTOK
//END BLEERN - let the system crash if we try to allocate too many handles!

	imul.ebx	ebx, sizeof (OneHandle)
	push		  edi
	l.edi		  #handlesrt					   // there is an compiler error
	add.ebx		edi							   // this is the reason wy we do this different
	pop			  edi

	s.ax		  (ebx+OneHandle.Typ)
	s.edi		  (ebx+OneHandle.thisp)

	test.ax		DmCallProg						// test if it is Main Prog
	jz			  getHandleRtSB
	add.ecx		StartOfRt
	add.ecx		offset
	s.cx		  (ebx+OneHandle.Address)
	l.eax		  ecx								// handle
	jmp			  getHandleRtMain

getHandleRTSB
	add.edx		StartOfCode
	add.edx		offset
	s.dx		  (ebx+OneHandle.Address)
	l.eax		  edx

getHandleRtMain

	inc.w		  HandleNrRT

GetHandleRet
	pop			  ecx
	pop			  edx

END_FUNCTION
#endif

FUNCTION AWL DiasMasterMain::GetProgPointer
#ifdef _LSL_TARGETARCH_X86

// it is in the cyclic

	l.ebx		PtrCY
	l.edx   IPSub
	l.ecx		IPMainCy
	test.AX		Dmrealtime
	jz			GetProgP_Cy

// it is in the Realtime
	l.ebx		PtrRT
	l.ecx		IPMainRT
GetProgP_Cy
#endif
END_FUNCTION
//
//
//  --> ax is mode byte (realtime or cyclic)
//		ECX = IP of the Mainprog
//		EDX = IP of the subprog
FUNCTION AWL DiasMasterMain::StoreNewPointers
#ifdef _LSL_TARGETARCH_X86
	s.edx		  IPSub
	and.ax		DmRealtime
	jnz			  StoreNewPRT		// --> realtime
	s.ecx		  IPMainCY
	jmp			  StoreNewRet

StoreNewPRT
	s.ecx		  IPMainRT
StoreNewRet
#endif
END_FUNCTION
// ****************************************
//   einmal das programm linken
// ****************************************
// the main and the subprogramms are linked together
// also the calls are linked with the absolute adresse
#ifdef _LSL_TARGETARCH_ARM
FUNCTION DiasMasterMain::LinkMaster
  VAR
  	pSINT : ^SINT;
  END_VAR

// ****************************************
//   add the "END" to the cyclic programm
// ****************************************

  (#CallsCY[0] + IPMainCY)^ := dbEnd;
  IPMainCY += 1;

// *******************************************************
//   add the "JMP to Begin" to the RT Programm
//   + mov timer to RAMCELL to calculate the right timing
// *******************************************************

  pSINT := #CallsRT[0] + IPMainRT;
  (pSINT + MovStruct.Opc)^        := dbMov;
  (pSINT$^UINT + MovStruct.Srce)^  := DmPllTmrAct;
  (pSINT$^UINT + MovStruct.Dest)^  := DmUserData;

  pSINT    += sizeof(MovStruct);
  IPMainRt += sizeof(MovStruct);

  ud_DelayRealtime += C_TimeMove;

  // Mark realtime task of intelligent master as inactive
  (pSINT + MovStruct.Opc)^        := dbMov;
  (pSINT$^UINT + MovStruct.Srce)^  := DmUserData + 2;
  (pSINT$^UINT + MovStruct.Dest)^  := DmUserData + 3;

  pSINT    += sizeof(MovStruct);
  IPMainRt += sizeof(MovStruct);

  ud_DelayRealtime += C_TimeMove;

  (pSINT + JmpStruct.Opc)^          := dbJmp;
  (pSINT$^UINT + JmpStruct.Adress)^  := StartOfRt$UINT;

  IPMainRT += sizeof(JmpStruct);

  ud_DelayRealtime += C_TimeJump;

END_FUNCTION
#else
FUNCTION AWL DiasMasterMain::LinkMaster
  VAR
    SizeofMainCY : DINT;
    SizeofMainRT : DINT;
  END_VAR

// ****************************************
//   add the "END" to the cyclic programm
// ****************************************

	l.ebx		  IPMainCy
	l.edi		  #CallsCY
	l.b			  (ebx+edi),dbend
	inc.d		  IPMainCy

// *******************************************************
//   add the "JMP to Begin" to the RT Programm
//   + mov timer to RAMCELL to calculate the right timing
// *******************************************************

	l.ebx		  IPMainRt
	l.edi		  #CallsRt

	l.b			  (ebx+edi+MovStruct.Opc),dbMov
	l.w			  (ebx+edi+MovStruct.Srce),DmPllTmrAct
	l.w			  (ebx+edi+MovStruct.Dest),DmUserData

	add.ebx		sizeof (MovStruct)
	add.d		  IPMainRT, sizeof (MovStruct)

	ADD.D		  ud_DelayRealtime,C_TimeMove		//#SR001

	//#SR010 start Mark realtime task of intelligent master as inactive
	l.b			  ( ebx + edi + MovStruct.Opc ), dbMov
	l.w			  ( ebx + edi + MovStruct.Srce ), DmUserData + 2
	l.w			  ( ebx + edi + MovStruct.Dest ), DmUserData + 3

	add.ebx		sizeof (MovStruct)
	add.d		  IPMainRT, sizeof (MovStruct)

	ADD.D		  ud_DelayRealtime,C_TimeMove
	//#SR010 end

	l.b			  (ebx+edi+JmpStruct.Opc),dbJmp
	l.eax		  startofrt
	s.ax		  (ebx+edi+JmpStruct.Adress)

	add.d		  IPMainRT, sizeof (JmpStruct)

	ADD.D		  ud_DelayRealtime,C_TimeJump		//#SR001

END_FUNCTION
#endif

// ********************************************************
//  .. load the cyclic programm in to the master
// ********************************************************
#ifdef _LSL_TARGETARCH_ARM
FUNCTION DiasMasterMain::LoadCyclicProg
  VAR
    Counter : DINT;
    pCalls  : ^USINT;
    pProg   : ^USINT;
    pUSINT  : ^USINT;
  END_VAR

  // with help variable we get only half of the ARM assembler code for the assignment
  pUSINT := _IOSEGMENT$^USINT + DmState;
  pUSINT^ := pUSINT^ AND 16#0F;   // all cyclic programs OFF

  pProg := _IOSEGMENT$^USINT + (_IOSEGMENT$^UINT + DmCyStartAdrM0)^;  // load start of program

  pCalls  := #CallsCY[0];
  Counter := IPMainCY + 1;

  while Counter do
    pProg^ := pCalls^;

    pCalls += 1;
    pProg += 1;
    Counter -= 1;
  end_while;

END_FUNCTION

#else
FUNCTION AWL DiasMasterMain::LoadCyclicProg

	L.EDI		  _IOSEGMENT
	L.AL		  (EDI+DmState)           // All Cyclic Programms OFF
	and.al		16#0f
	S.AL		  (EDI+DmState)

	clr			  ebx
	L.BX		  (EDI+DmCyStartAdrM0)      // load start of programm

	l.edx		  #CallsCY
	l.ecx		  IPMainCY
	inc			  ecx

LoadCyLoop
	l.al		  (edx)
	s.al		  (ebx+edi)
	inc			  ebx
	inc			  edx
	loop		  LoadCyLoop

END_FUNCTION
#endif

#ifdef _LSL_TARGETARCH_ARM
FUNCTION DiasMasterMain::StartCyclicProg
  VAR
  	pUSINT  : ^USINT;
  END_VAR

  // with help variable we get only half of the ARM assembler code
  pUSINT := _IOSEGMENT$^USINT + DmState;

  // Cyclic Programms ON Master 1
  pUSINT^ := pUSINT^ OR 16#10;

END_FUNCTION
#else
FUNCTION AWL DiasMasterMain::StartCyclicProg

	L.EDI		_IOSEGMENT
	L.AL		(EDI+DmState)           // Cyclic Programms ON Master 1
	OR.AL		16#10
	S.AL		(EDI+DmState)

END_FUNCTION
#endif

#ifdef _LSL_TARGETARCH_ARM
FUNCTION DiasMasterMain::StartRealtimeProg
  VAR
  	pUSINT  : ^USINT;
  END_VAR

  // with help variable we get only half of the ARM assembler code
  pUSINT := _IOSEGMENT$^USINT + DmState;

  // Realtime Programms ON Master 1
  pUSINT^ := pUSINT^ OR 16#01;

END_FUNCTION
#else
FUNCTION AWL DiasMasterMain::StartRealtimeProg

	L.EDI		_IOSEGMENT
	L.AL		(EDI+DmState)           // Cyclic Programms ON Master 1
	OR.AL		16#01
	S.AL		(EDI+DmState)

END_FUNCTION
#endif

// ********************************************************
//  .. load the cyclic programm into the master
// ********************************************************
FUNCTION DiasMasterMain::LoadRealtimeProg
  VAR
    Counter : DINT;
    pCalls  : ^USINT;
    pProg   : ^USINT;
    pUSINT  : ^USINT;
  END_VAR

  // with help variable we get only half of the ARM assembler code for the assignment
  pUSINT := _IOSEGMENT$^USINT + DmState;
  pUSINT^ := pUSINT^ AND 16#F0;   // all realtime programs OFF

  pProg := _IOSEGMENT$^USINT + (_IOSEGMENT$^UINT + DmRtStartAdrM0)^;  // load start of program

  pCalls  := #CallsRT[0];
  Counter := IPMainRT + 1;

  while Counter do
    pProg^ := pCalls^;

    pCalls += 1;
    pProg += 1;
    Counter -= 1;
  end_while;

END_FUNCTION

FUNCTION  DiasMasterMain::CallUpdata
  VAR_INPUT
    Thisp		  : pHwBase;
    Handle		: UDINT;
  END_VAR

	thisp^.updatecy(handle);

END_FUNCTION
FUNCTION  DiasMasterMain::CallUpdataRT
  VAR_INPUT
    Thisp		  : pHwBase;
    Handle		: UDINT;
  END_VAR

	thisp^.updatert(handle);

END_FUNCTION

//[#ENGLISH]
//0= connected direct to master
//1= connected via CIC
//
//
//-1 = fault
FUNCTION VIRTUAL GLOBAL DiasMasterMain::GetConnection
  VAR_OUTPUT
    CType		: DINT;
  END_VAR

	CType :=0;		// we are the main controller

END_FUNCTION

//[#ENGLISH]
//read one Byte from C-DIAS bus on Board
#pragma warning (disable:73)
FUNCTION VIRTUAL GLOBAL DiasMasterMain::I2CReadOneByte
  VAR_INPUT
    AdressCDIAS	: UINT;
    pData		    : ^USINT;
  END_VAR
  VAR_OUTPUT
    result		  : DINT;
  END_VAR

	result:=-1;

END_FUNCTION
#pragma warning (default:73)

FUNCTION VIRTUAL GLOBAL DiasMasterMain::GetEEState
  VAR_OUTPUT
    State		: DINT;
  END_VAR

	State := CDiasType;

END_FUNCTION

#pragma warning (disable:73)
FUNCTION VIRTUAL GLOBAL DiasMasterMain::ReadEEData
  VAR_INPUT
    Adress		: UDINT;
    pData		  : ^USINT;
  END_VAR
  VAR_OUTPUT
    retval		: DINT;
  END_VAR

	retval := -1;

END_FUNCTION
#pragma warning (default:73)

#ifdef _LSL_TARGETARCH_ARM
FUNCTION VIRTUAL GLOBAL DiasMasterMain::AddCall2List
  VAR_INPUT
    Mode		    : UINT;
    RTCY		    : DINT;
    thisp		    : ^void;
    callOptions : USINT;
  END_VAR
  VAR_OUTPUT
    Handle		  : DINT;
  END_VAR

  if (RTCY AND DmRealtime) = DmRealtime then
    ARM_EAX := RTCY$UDINT OR DmCallProg;
    ARM_EDI := thisp$UDINT;
    GetHandle(HandleNrRT, callOptions);
    Handle := ARM_EAX$DINT;
  else
    ARM_EAX := RTCY$UDINT OR DmCallProg;
    ARM_EDI := thisp$UDINT;
    GetHandle(HandleNrCY, callOptions);
    Handle := ARM_EAX$DINT;
  end_if;

END_FUNCTION

#else

FUNCTION AWL VIRTUAL GLOBAL DiasMasterMain::AddCall2List
	VAR_INPUT
		Mode 	      : UINT;
		RTCY 	      : DINT;
		thisp 	    : ^void;
		callOptions : USINT;
	END_VAR
	VAR_OUTPUT
		Handle 	    : DINT;
	END_VAR

	l.ecx		  16#8000					//Because we got equal handles and ecx register wasn't set //#SR000

	l.ax		  RTCY+0
	or.ax		  DmCallProg				// this is in the Main
	l.edi		  thisp

    // changed not CallStruct.Mode because we need for each add call a different number
    // and therefore we take IP off programm

	test.ax		Dmrealtime
	jnz			  AddCall2ListRT
	lzxw.ebx	HandleNrCY
	jmp			  AddCall2ListCy
AddCall2ListRT
	lzxw.ebx	HandleNrRT
AddCall2ListCy

  push.b    callOptions

	push		  ebx
	call		  GetHandle
  add.esp   5
	s.eax		  handle

END_FUNCTION
#endif

#ifdef _LSL_TARGETARCH_ARM
FUNCTION VIRTUAL GLOBAL DiasMasterMain::CyWorkStdMas
  VAR
#ifdef TRIGGER_WD_386_IN_CYCLIC
    TempAL    : SINT;
#endif
    TempEBX   : DINT;
    i         : UDINT;
    pHandle   : ^OneHandle;
  //-------------------------------------Profiler Start----------------------------------------------
#ifdef DiasMasterC_Profiler
    MuSecTime : UDINT;
  END_VAR

  MuSecTime := OS_ReadMicroSec();
  //Anfangsdelay abwarten
	if MuSecTime - DMC_Time_CY.init > DM_ProfilerDelay then
    DMC_Time_CY.start  := MuSecTime;    //Startzeit nehmen
    DMC_Time_CY.initfl := FALSE;        //Initflag löschen
  else
    DMC_Time_CY.initfl := TRUE;         //Initflag setzen
  end_if;
//-------------------------------------Profiler End------------------------------------------------
#else
  END_VAR
#endif

  WriteRTLogs();

  if ops.tAbsolute <> OldTime then

#ifdef TRIGGER_WD_386_IN_CYCLIC
// ** hier mal den watchdog triggern ** #FA  (Watchdog der CCL)
//ist interner CPU Watchdog --> kein Abfall der Hardware wenn nicht getriggert wird

    if (_WhoAmI = 16#23) |  (_WhoAmI = 16#27) | (_WhoAmI = 16#28) | (_WhoAmI = 16#29) then
      if _RTOSVersion >= OSVersionDIASIO then
	//*****************************************************
	//***** use OS functions instead of own functions *****
	//*****************************************************
        CCLWatchdog_Trigger();
      else
	//*****************************************************
	//*** use own functions (should be obsolete by now) ***
	//*****************************************************
        TraceAsyncError();
      end_if;
    end_if;
#endif

// **************************************************
//  now take data and call update function with thisp
// **************************************************
    CyclicReady := TRUE;

    if HandleNrCy then
      pHandle := #HandlesCY[0];

      for i := 0 to HandleNrCy-1 do
        if pHandle^.Typ AND DmCallProg then
          pHandle^.thisp^.UpdateCy(pHandle^.Address);
        end_if;

        pHandle += sizeof(OneHandle);
      end_for;
    end_if;

    if _RTOSVersion >= OSVersionDIASIO then
	//*****************************************************
	//***** use OS functions instead of own functions *****
	//*****************************************************
      UpdateRetryCounter();
    else
	//*****************************************************
	//*** use own functions (should be obsolete by now) ***
	//*****************************************************
      if (_WhoAmI = 16#17) | (_WhoAmI = 16#19) then
        UpdateRetryCounter();
      else
        if _IOSegment then
          if _IOSegment = 16#D0000 then
            TraceAsyncError();
          else
            TempEBX := to_DINT((_IOSegment$^SINT + 16#C008)^);
          end_if;

          DIASRetryCounter += TempEBX$USINT - oldErrorCounter$USINT;
          oldErrorCounter := TempEBX;
        end_if;
      end_if;
    end_if;
  end_if;
  OldTime := ops.tAbsolute;

  // look if we got the pointer to the safety manager
  if SafetyManagerThis then
    // call safety manager
    SafetyManagerThis^.CyWork(0);
  end_if;

//-------------------------------------Profiler Start----------------------------------------------
#ifdef DiasMasterC_Profiler
  //schaun ob Delayzeit schon abgelaufen ist
  if DMC_Time_CY.initfl = FALSE then
    MuSecTime := OS_ReadMicroSec();

    DMC_Time_CY.stop := MuSecTime;        //Stopzeit speichern

    MuSecTime -= DMC_Time_CY.start;       //Differenz berechnen
    MuSecTime -= DM_CPUconstant;          //Zeit für OS_REadMicroSec - Funktion subtrahieren

    DMC_Time_CY.diff := MuSecTime;        //korr. Differenz speichern
    DMC_Time_CY.sum  += MuSecTime;        //Zur Summe addieren

    DMC_Time_CY.run  += 1;                //Durchlaufzähler erhöhen

    if MuSecTime < DMC_Time_CY._min then
      DMC_Time_CY._min := MuSecTime;      //Minimalzeit speichern
    end_if;

    if MuSecTime > DMC_Time_CY._max then
      DMC_Time_CY._max := MuSecTime;      //Maximalzeit speichern
    end_if;

    //Durchschnitt berechnen
    //*100 damit wir 2 Kommastellen haben
    DMC_Time_CY.avg := DMC_Time_CY.sum * 100 / DMC_Time_CY.run;
  end_if;

#endif
//-------------------------------------Profiler End------------------------------------------------

END_FUNCTION

#else

FUNCTION AWL VIRTUAL GLOBAL DiasMasterMain::CyWorkStdMas

//#wp001
//============================ Profiler start======================================================
#ifdef  DiasMasterC_Profiler
	CLI											//damit keine Interrupts die Messung stören
	push 		  edi
	push 		  eax
	l.edi 		_LSL_POS
	l.edi 		( edi + DM_LSLPOS_SYSTIME )
	l.edi 		( edi + DM_LSLSYSTIME_MICROSEC )
	call		  edi								//OS_ReadMicroSec - Funktion aufrufen
	l.ebx		  eax
	sub.ebx		DMC_Time_CY.init					//Anfangsdelay abwarten
	cmp.ebx		DM_ProfilerDelay
	jle			  LABEL_DMCPREEND
	s.eax 		DMC_Time_CY.start					//Startzeit nehmen
	x.cl		  cl
	s.cl		  DMC_Time_CY.initfl				//Initflag löschen
	jmp 		  LABEL_DMCstartfunc

LABEL_DMCPREEND
	l.b		    DMC_Time_CY.initfl,1					//Initflag setzen

LABEL_DMCstartfunc
	pop 		  eax
	pop 		  edi
#endif
//============================ Profiler end========================================================

  cmp.b     SkipCy,1
  je        NoLocalSafety2

	l.eax		  OPS.Tabsolute
	cmp.eax		oldtime
	je			  NoCyclProgEnd // #BS003
	s.eax		  oldtime

#ifdef TRIGGER_WD_386_IN_CYCLIC

// ** hier mal den watchdog triggern ** #FA  (Watchdog der CCL)
//ist interner CPU Watchdog --> kein Abfall der Hardware wenn nicht getriggert wird

 	CMP.D		  _WhoAmI,16#23 // #BS003

	//#SR002 Start
	je			  CCLWatchdog
	cmp.d		  _WhoAmI,16#27
	je			  CCLWatchdog
	cmp.d		  _WhoAmI,16#28
	je			  CCLWatchdog
	cmp.d		  _WhoAmI,16#29
	jne			  NoCCLWatchdog

CCLWatchdog
	//#SR002 End

	//ws005
	//*****************************************************
	//***** use OS functions instead of own functions *****
	//*****************************************************
	cmp.d		  _RTOSVersion, OSVersionDIASIO
	jl			  LABEL_OLDWD
  call    	CCLWatchdog_Trigger
	jmp			  NoCCLWatchdog

LABEL_OLDWD
	//*****************************************************
	//*** use own functions (should be obsolete by now) ***
	//*****************************************************
	// /ws005

	l.dx		  16#f862
	inb
	or			  16#40
	outb
	and			  2#10111111
	outb
	// /ws005

NoCCLWatchdog
#endif

// **************************************************
//  now take data and call update function with thisp
// **************************************************
	l.b 		  CyclicReady,1	//ws005

	l.ebx		  #HandlesCY
	lzxw.ecx	HandleNrCy
	jecxz		  NoCyclProg

HandleLoop
	test.w		(ebx+OneHandle.Typ),DmCallProg
	jz			  NextHandle

	push		  ecx
	push		  ebx

	L.eax		  (ebx+OneHandle.thisp)
	LZXW.ECX	(ebx+OneHandle.Address)
	push		  ecx
	push		  eax
	call		  CallUpdata
	add.esp		8

	pop			  ebx
	pop			  ecx

NextHandle
	add.ebx		sizeof (OneHandle)
	loop		  HandleLoop
NoCyclProg

//ws004

	//ws005
	//*****************************************************
	//***** use OS functions instead of own functions *****
	//*****************************************************
	cmp.d		  _RTOSVersion, OSVersionDIASIO
	jl			  LABEL_OLDUPDATE
  call      UpdateRetryCounter	// this function will also run with ETT321 and ET261
	jmp			  NoCyclProgEND

LABEL_OLDUPDATE
	//*****************************************************
	//*** use own functions (should be obsolete by now) ***
	//*****************************************************
	cmp.d		  _WHOAMI, 16#19
	je			  LABEL_ET2XX
	cmp.d		  _WHOAMI, 16#17
	je			  LABEL_ET2XX
	jmp			  LABEL_CONT

LABEL_ET2XX
	call      UpdateRetryCounter	// this function will also run with ETT321 and ET261
	jmp		    NoCyclProgEND

LABEL_CONT
	// /ws005

// #BS003 Start
// #BS007 Start
	L.EDI		  _IOSegment
	//#SR019 start				//if _IOSegment = 0 we do not update retry counter
	o.edi		  edi
	jz			  NoCyclProgEND
	//#SR019 end

	CMP.EDI		16#D0000
	JNE			  Retry386
	PUSHF
	CLI

	l.dx		  16#335
	l			    1 // switch to control
	outb

	LZXB.EBX	(edi+16#4008)

	l.dx		  16#335
	clr			  al
	outb

	POPF
	JMP			  UpdateCount
Retry386
	Lzxb.ebx	(EDI+16#C008)

UpdateCount
// #BS007 End
	l.eax		  oldErrorCounter
	s.ebx		  oldErrorCounter
// #BS016 Start
	sub.bl		al
	lzxb.ebx	bl
	add.d		  DIASRetryCounter,eBx
NoCyclProgEND
// #BS003 End

  // look if we got the pointer to the safety manager
  cmp.d     SafetyManagerThis, 0
  je        NoLocalSafety2

  // call safety manager
  CALL      CallSafetyManager

NoLocalSafety2

//#wp001
//============================ Profiler end======================================================
#ifdef  DiasMasterC_Profiler
	cmp.b 		DMC_Time_CY.initfl, 1				//schaun ob Delayzeit schon abgelaufen ist
	je			  LABEL_DMCEND
	pushad
	l.edi 		_LSL_POS
	l.edi 		( edi + DM_LSLPOS_SYSTIME )
	l.edi 		( edi + DM_LSLSYSTIME_MICROSEC )
	call		  edi								//OS_REadMicroSec - Funktion aufrufen
	s.eax 		DMC_Time_CY.stop					//Stopzeit speichern
	l.ebx 		DMC_Time_CY.start
	sub.eax		ebx								//Differenz berechnen
	sub.eax		DM_CPUconstant					//Zeit für OS_REadMicroSec - Funktion subtrahieren
	s.eax 		DMC_Time_CY.diff					//Ergebnis speicern
	l.ebx 		DMC_Time_CY.sum
	add.ebx 	eax								//Zur Summe addieren
	s.ebx 		DMC_Time_CY.sum					//Summe speichern
	l.ecx		  DMC_Time_CY.run
	inc 		  ecx								//Durchlaufzähler erhöhen
	s.ecx 		DMC_Time_CY.run					//Durchlaufzähler speichern
	cmp.eax		DMC_Time_CY._min					//mit Minimalzeit vergleichen
	jae			  LABEL_DMCcont
	s.eax 		DMC_Time_CY._min					//Minimalzeit speichern

LABEL_DMCcont
	cmp.eax 	DMC_Time_CY._max					//Mit Maximalzeit vergleichen
	jbe 		  LABEL_DMCcont1
	s.eax 		DMC_Time_CY._max					//Maximalzeit speichern

LABEL_DMCcont1
	l.eax		  ebx								//Summe in al laden
	imul.eax	eax,100							//*100 damit wir 2 Kommastellen haben
	x.edx 		edx
	idiv		  ecx								//durch Durchläufe dividieren
	s.eax		  DMC_Time_CY.avg					//Durchschnitt speichern
	popad

LABEL_DMCEND
	STI
#endif
//============================ Profiler end========================================================

END_FUNCTION
#endif

#ifdef _LSL_TARGETARCH_ARM
FUNCTION VIRTUAL GLOBAL DiasMasterMain::RtWorkStdMas
#ifdef DM_DEBUG_ARM
  // This method is not supported with ARM
  ((0)$^USINT)^ := 0;
#endif
END_FUNCTION
#else
FUNCTION AWL VIRTUAL GLOBAL DiasMasterMain::RtWorkStdMas

//#wp001
//============================ Profiler start======================================================
#ifdef  DiasMasterC_Profiler
	CLI											//damit keine Interrupts die Messung stören
	push 		  edi
	push 		  eax
	l.edi 		_LSL_POS
	l.edi 		( edi + DM_LSLPOS_SYSTIME )
	l.edi 		( edi + DM_LSLSYSTIME_MICROSEC )
	call		  edi								//OS_ReadMicroSec - Funktion aufrufen
	l.ebx		  eax
	sub.ebx		DMC_Time_RT.init					//Anfangsdelay abwarten
	cmp.ebx		DM_ProfilerDelay
	jle			  LABEL_DMCPREEND
	s.eax 		DMC_Time_RT.start					//Startzeit nehmen
	x.cl		  cl
	s.cl		  DMC_Time_RT.initfl				//Initflag löschen
	jmp 		  LABEL_DMCstartfunc

LABEL_DMCPREEND
	l.b		    DMC_Time_RT.initfl,1					//Initflag setzen

LABEL_DMCstartfunc
	pop 		  eax
	pop 		  edi
#endif
//============================ Profiler end========================================================
  cmp.b			b_PllInit, TRUE
	je				LABEL_NoStart

	//in first run we start pll
	call			StartPll
	l.b				b_PllInit, TRUE
LABEL_NoStart

#ifndef TRIGGER_WD_386_IN_CYCLIC

// ** hier mal den watchdog triggern ** #FA  (Watchdog der CCL)
//ist interner CPU Watchdog --> kein Abfall der Hardware wenn nicht getriggert wird

 	CMP.D		  _WhoAmI,16#23 // #BS003

	//#SR002 Start
	je			  CCLWatchdog
	cmp.d		  _WhoAmI,16#27
	je			  CCLWatchdog
	cmp.d		  _WhoAmI,16#28
	je			  CCLWatchdog
	cmp.d		  _WhoAmI,16#29
	je			  CCLWatchdog
	cmp.d		  _WhoAmI,16#35
	je			  CCLWatchdog
	cmp.d		  _WhoAmI,16#34
	jne			  NoCCLWatchdog

CCLWatchdog
	//#SR002 End

	//ws005
	//*****************************************************
	//***** use OS functions instead of own functions *****
	//*****************************************************
	cmp.d		  _RTOSVersion, OSVersionDIASIO
	jl			  LABEL_OLDWD
  	call   	CCLWatchdog_Trigger
	jmp			  NoCCLWatchdog

LABEL_OLDWD
	//*****************************************************
	//*** use own functions (should be obsolete by now) ***
	//*****************************************************
	// /ws005

	l.dx		  16#f862
	inb
	or			  16#40
	outb
	and			  2#10111111
	outb
	// /ws005

NoCCLWatchdog
#endif

#IFNDEF OldDiasXilinx // global sync
	l.ebx		  RTBSyncAdr
	o.ebx		  ebx
	jz			  RtNoRTB
	//ws005
	//*****************************************************
	//***** use OS functions instead of own functions *****
	//*****************************************************
	cmp.d		  _RTOSVersion, OSVersionDIASIO
	jl			  LABEL_MAYBEOLDUPDATE
	push.d		0     //data to write
	push.d		2     //offset
	push.d		63    //DIAS place
	l.eax		  pDIAS
	push		  eax   //DIAS structure
	call		  ( eax + 27 )  //call to OS function OS_DIAS_WriteCtrl_
	add.esp		16
	jmp			  RtNoRTB

LABEL_MAYBEOLDUPDATE
	cmp.d		  _WHOAMI, 16#19
	je			  LABEL_ISETXX
	cmp.d		  _WHOAMI, 16#17
	jne			  LABEL_OLDUPDATE

LABEL_ISETXX
	push.d		0     //data to write
	push.d		2     //offset
	push.d		63    //DIAS place
	l.eax		  pDIAS
	push		  eax   //DIAS structure
	call		  ( eax + 27 )  //call to OS function OS_DIAS_WriteCtrl_
	add.esp		16
	jmp			  RtNoRTB

LABEL_OLDUPDATE
  l.edi		  _ioSegment  //ws005
	s			    ( ebx + edi )

	// /ws005

#ELSE // local sync
	LZXB.ECX	NumberSyncs
	JECXZ		  RtNoRTB

	L.EDX		  #RtbLocalSyncAdr[0]
SyncJMP
	l.edi		  _ioSegment  //ws005
	LZXW.EBX	(EDX)
	L.B			  (ebx+edi),1
	ADD.EDX		SIZEOF(HINT)
	LOOP		  SyncJMP
#ENDIF

RtNoRTB
// **************************************************
//  now take data and call update function with thisp
// **************************************************
	l.b			  RealtimeReady,1		//ws005

	l.ebx		  #HandlesRt
	lzxw.ecx	HandleNrRt
	jecxz		  LABEL_RtPostScan

HandleLoopRt
	test.w		(ebx+OneHandle.Typ),DmCallProg
	jz			  NextHandleRt

	push		  ecx
	push		  ebx

	L.eax		  (ebx+OneHandle.thisp)
	LZXW.ECX	(ebx+OneHandle.Address)
	push		  ecx
	push		  eax

	call		  CallUpdataRT
	add.esp		8

	pop			  ebx
	pop			  ecx

NextHandleRt
	add.ebx		sizeof (OneHandle)
	loop		  HandleLoopRt

LABEL_RtPostScan

//BLEERN START
  cmp.d     HwControl, 0
  jne       NoRtProg

  call      UpdateRtPostScan
//BLEERN ENDE

NoRtProg

	FC			WDDIAS

//#wp001
//============================ Profiler end======================================================
#ifdef  DiasMasterC_Profiler
	cmp.b 		DMC_Time_RT.initfl, 1				//schaun ob Delayzeit schon abgelaufen ist
	je			  LABEL_DMCEND
	pushad
	l.edi 		_LSL_POS
	l.edi 		( edi + DM_LSLPOS_SYSTIME )
	l.edi 		( edi + DM_LSLSYSTIME_MICROSEC )
	call		  edi								//OS_REadMicroSec - Funktion aufrufen
	s.eax 		DMC_Time_RT.stop					//Stopzeit speichern
	l.ebx 		DMC_Time_RT.start
	sub.eax		ebx								//Differenz berechnen
	sub.eax		DM_CPUconstant					//Zeit für OS_REadMicroSec - Funktion subtrahieren
	s.eax 		DMC_Time_RT.diff					//Ergebnis speicern
	l.ebx 		DMC_Time_RT.sum
	add.ebx 	eax								//Zur Summe addieren
	s.ebx 		DMC_Time_RT.sum					//Summe speichern
	l.ecx		  DMC_Time_RT.run
	inc 		  ecx								//Durchlaufzähler erhöhen
	s.ecx 		DMC_Time_RT.run					//Durchlaufzähler speichern
	cmp.eax		DMC_Time_RT._min					//mit Minimalzeit vergleichen
	jae			  LABEL_DMCcont
	s.eax 		DMC_Time_RT._min					//Minimalzeit speichern

LABEL_DMCcont
	cmp.eax 	DMC_Time_RT._max					//Mit Maximalzeit vergleichen
	jbe 		  LABEL_DMCcont1
	s.eax 		DMC_Time_RT._max					//Maximalzeit speichern

LABEL_DMCcont1
	l.eax		  ebx								//Summe in al laden
	imul.eax	eax,100							//*100 damit wir 2 Kommastellen haben
	x.edx 		edx
	idiv		  ecx								//durch Durchläufe dividieren
	s.eax		  DMC_Time_RT.avg					//Durchschnitt speichern
	popad

LABEL_DMCEND
	STI
#endif
//============================ Profiler end========================================================

END_FUNCTION
#endif

FUNCTION VIRTUAL GLOBAL DiasMasterMain::GetMasterType
  VAR_OUTPUT
    MasterType		: UDINT;
  END_VAR

  MasterType:=DiasType;

END_FUNCTION

FUNCTION VIRTUAL GLOBAL DiasMasterMain::GetCDiasIosegment
  VAR_OUTPUT
    CIOSegment		: ^USINT;
  END_VAR

  CIOSegment := CDiasHwPointer;

END_FUNCTION

#ifdef _LSL_TARGETARCH_ARM
FUNCTION VIRTUAL GLOBAL DiasMasterMain::RtWorkStdMasIPC
#ifdef _LSL_TARGETARCH_X86
  VAR
    i         : DINT;
    pHandle   : ^OneHandle;
  #ifdef OldDiasXilinx
    pHINT     : ^HINT;
  #endif
  //-------------------------------------Profiler Start----------------------------------------------
  #ifdef DiasMasterC_Profiler
    MuSecTime : UDINT;
  END_VAR

  MuSecTime := OS_ReadMicroSec();
  //Anfangsdelay abwarten
	if MuSecTime - DMC_Time_RT.init > DM_ProfilerDelay then
    DMC_Time_RT.start  := MuSecTime;    //Startzeit nehmen
    DMC_Time_RT.initfl := FALSE;        //Initflag löschen
  else
    DMC_Time_RT.initfl := TRUE;         //Initflag setzen
  end_if;
//-------------------------------------Profiler End------------------------------------------------
#else
  END_VAR
#endif

#IFNDEF OldDiasXilinx // global sync
  if RTBSyncAdr then
    CLI();

    To_OSKernel.OutByte(Portnumber:=16#335, value:=1);

    (_IOSegment$^USINT + RTBSyncAdr$UDINT - 16#8000)^ := 1;

    To_OSKernel.OutByte(Portnumber:=16#335, value:=0);

    STI();
  end_if;
#ELSE // local sync
  if NumberSyncs then
    CLI();

    To_OSKernel.OutByte(Portnumber:=16#335, value:=1);

    pHINT := #RtbLocalSyncAdr[0];
    for i := 0 to NumberSyncs-1 do
      (_IOSegment$^SINT + pHINT^ - 16#8000)^ := 1;

      pHINT += sizeof(HINT);
    end_for;

    To_OSKernel.OutByte(Portnumber:=16#335, value:=0);

    STI();
  end_if;
#ENDIF

// **************************************************
//  now take data and call update function with thisp
// **************************************************
  RealtimeReady := 1;

  // call update methods with thispointer
  if HandleNrRt then
    pHandle := #HandlesRT[0];
    for i := 0 to HandleNrRT-1 do
      if pHandle^.Typ AND DmCallProg then
        pHandle^.thisp^.UpdateRt(pHandle^.Address);
      end_if;

      pHandle += sizeof(OneHandle);
    end_for;
  end_if;

  if HwControl = 0 then
    UpdateRtPostScan();
  end_if;

  WDDIAS();

//-------------------------------------Profiler Start----------------------------------------------
#ifdef DiasMasterC_Profiler
  //schaun ob Delayzeit schon abgelaufen ist
  if DMC_Time_RT.initfl = FALSE then
    MuSecTime := OS_ReadMicroSec();

    DMC_Time_RT.stop := MuSecTime;        //Stopzeit speichern

    MuSecTime -= DMC_Time_RT.start;       //Differenz berechnen
    MuSecTime -= DM_CPUconstant;          //Zeit für OS_REadMicroSec - Funktion subtrahieren

    DMC_Time_RT.diff := MuSecTime;        //korr. Differenz speichern
    DMC_Time_RT.sum  += MuSecTime;        //Zur Summe addieren

    DMC_Time_RT.run  += 1;                //Durchlaufzähler erhöhen

    if MuSecTime < DMC_Time_RT._min then
      DMC_Time_RT._min := MuSecTime;      //Minimalzeit speichern
    end_if;

    if MuSecTime > DMC_Time_RT._max then
      DMC_Time_RT._max := MuSecTime;      //Maximalzeit speichern
    end_if;

    //Durchschnitt berechnen
    //*100 damit wir 2 Kommastellen haben
    DMC_Time_RT.avg := DMC_Time_RT.sum * 100 / DMC_Time_RT.run;
  end_if;

#endif
//-------------------------------------Profiler End------------------------------------------------
#endif
END_FUNCTION
#else
FUNCTION AWL VIRTUAL GLOBAL DiasMasterMain::RtWorkStdMasIPC

//#wp001
//============================ Profiler start======================================================
#ifdef  DiasMasterC_Profiler
	CLI											//damit keine Interrupts die Messung stören
	push 		  edi
	push 		  eax
	l.edi 		_LSL_POS
	l.edi 		( edi + DM_LSLPOS_SYSTIME )
	l.edi 		( edi + DM_LSLSYSTIME_MICROSEC )
	call		  edi								//OS_ReadMicroSec - Funktion aufrufen
	l.ebx		  eax
	sub.ebx		DMC_Time_RT.init					//Anfangsdelay abwarten
	cmp.ebx		DM_ProfilerDelay
	jle			  LABEL_DMCPREEND
	s.eax 		DMC_Time_RT.start					//Startzeit nehmen
	x.cl		  cl
	s.cl		  DMC_Time_RT.initfl				//Initflag löschen
	jmp 		  LABEL_DMCstartfunc

LABEL_DMCPREEND
	l.b		    DMC_Time_RT.initfl,1					//Initflag setzen

LABEL_DMCstartfunc
	pop 		  eax
	pop 		  edi
#endif
//============================ Profiler end========================================================

	l.edi		  _ioSegment

#IFNDEF OldDiasXilinx // global sync
	l.ebx		  RTBSyncAdr
	o.ebx		  ebx
	jz			  RtNoRTB

	cli
	l.dx		  16#335
	l			    1
	outb
	sub.ebx		16#8000
	s			    (ebx+edi)
	clr			  al
	outb
	sti

#ELSE // local sync
	LZXB.ECX	NumberSyncs
	JECXZ		  RtNoRTB

	cli
	l.dx		  16#335
	l			    1 // switch to control
	outb

	L.EDX		  #RtbLocalSyncAdr[0]
SyncJMP
	LZXW.EBX	(EDX)

	sub.ebx		16#8000
	L.B			  (ebx+edi),1

	ADD.EDX		SIZEOF(HINT)
	LOOP		  SyncJMP

	l.dx		  16#335
	clr			  al
	outb
	sti

#ENDIF

RtNoRTB
// **************************************************
//  now take data and call update function with thisp
// **************************************************
	l.b			  RealtimeReady,1		//ws005

	l.ebx		  #HandlesRt
	lzxw.ecx	HandleNrRt
	jecxz		  LABEL_RtPostScan

HandleLoopRt
	test.w		(ebx+OneHandle.Typ),DmCallProg
	jz			  NextHandleRt

	push		  ecx
	push		  ebx

	L.eax		  (ebx+OneHandle.thisp)
	LZXW.ECX	(ebx+OneHandle.Address)
	push		  ecx
	push		  eax

	call		  CallUpdataRT
	add.esp		8

	pop			  ebx
	pop			  ecx

NextHandleRt
	add.ebx		sizeof (OneHandle)
	loop		  HandleLoopRt

LABEL_RtPostScan
//BLEERN START
  cmp.d     HwControl, 0
  jne       NoRtProg

  call      UpdateRtPostScan
//BLEERN ENDE

NoRtProg

	FC			  WDDIAS

//#wp001
//============================ Profiler end======================================================
#ifdef  DiasMasterC_Profiler
	cmp.b 		DMC_Time_RT.initfl, 1				//schaun ob Delayzeit schon abgelaufen ist
	je			  LABEL_DMCEND
	pushad
	l.edi 		_LSL_POS
	l.edi 		( edi + DM_LSLPOS_SYSTIME )
	l.edi 		( edi + DM_LSLSYSTIME_MICROSEC )
	call		  edi								//OS_REadMicroSec - Funktion aufrufen
	s.eax 		DMC_Time_RT.stop					//Stopzeit speichern
	l.ebx 		DMC_Time_RT.start
	sub.eax		ebx								//Differenz berechnen
	sub.eax		DM_CPUconstant					//Zeit für OS_REadMicroSec - Funktion subtrahieren
	s.eax 		DMC_Time_RT.diff					//Ergebnis speicern
	l.ebx 		DMC_Time_RT.sum
	add.ebx 	eax								//Zur Summe addieren
	s.ebx 		DMC_Time_RT.sum					//Summe speichern
	l.ecx		  DMC_Time_RT.run
	inc 		  ecx								//Durchlaufzähler erhöhen
	s.ecx 		DMC_Time_RT.run					//Durchlaufzähler speichern
	cmp.eax		DMC_Time_RT._min					//mit Minimalzeit vergleichen
	jae			  LABEL_DMCcont
	s.eax 		DMC_Time_RT._min					//Minimalzeit speichern

LABEL_DMCcont
	cmp.eax 	DMC_Time_RT._max					//Mit Maximalzeit vergleichen
	jbe 		  LABEL_DMCcont1
	s.eax 		DMC_Time_RT._max					//Maximalzeit speichern

LABEL_DMCcont1
	l.eax		  ebx								//Summe in al laden
	imul.eax	eax,100							//*100 damit wir 2 Kommastellen haben
	x.edx 		edx
	idiv		  ecx								//durch Durchläufe dividieren
	s.eax		  DMC_Time_RT.avg					//Durchschnitt speichern
	popad

LABEL_DMCEND
	STI
#endif
//============================ Profiler end========================================================

END_FUNCTION
#endif

FUNCTION  DiasMasterMain::WdCDIAS

  IF RTSSW <> 4 THEN
	  	//--- do watchdog while synchronizing -------------------
		#IFNDEF MaxWatchdog	// #BS016
		IF ops.tAbsolute - timestampCDIAS$UDINT > 100ms | RtDebug = 1 THEN			//#SR011
			timestampCDIAS$UDINT := ops.tAbsolute;
		#ENDIF

		//**** C - Dias Watchdog ****************************
			// #BS000
			IF (CDiasI2CWatchdog+2)^ AND 1 & MasterOn = 1 THEN // watchdogstatus (Bit0 = 1 => watchdog)
        bdRTLogs.Bit5 := 1;   //set Flag for Error Log
				MasterOn := 0;
				IMOFF := 1;
			ELSE
				IF MasterOn THEN
					CDiasI2CWatchdog^ := 0; // trigger watchdog
					// #BS002 only one watchdogregister for CDIAS and DIAS (IM)
				END_IF;
			END_IF;

			//**** Dias - Watchdog ******************************
			IF FirstModulFound <> 16#ff THEN		//ws005
				ReadKenn(FirstModulFound);
			END_IF;

		#IFNDEF MaxWatchdog	// #BS016
		END_IF;
		#ENDIF
  ELSE        //ws005: there is no point in triggering the WD twice while synchronizing

	#IFNDEF MaxWatchdog	// #BS016
    IF ops.tAbsolute - timestampCDIAS$UDINT > 100ms | RtDebug = 1 THEN			//#SR011
      timestampCDIAS$UDINT := ops.tAbsolute;
    #ENDIF
      //----- Always do CDIAS watchdog --------------------
      //**** C - Dias Watchdog *********************************************
      // #BS000
      IF (CDiasI2CWatchdog+2)^ AND 1 & MasterOn = 1 THEN // watchdogstatus (Bit0 = 1 => watchdog)
        bdRTLogs.Bit5 := 1;   //set Flag for Error Log
        MasterOn := 0;
        IMOFF := 1;
      ELSE
        IF MasterOn THEN
          CDiasI2CWatchdog^ := 0; // trigger watchdog
          // #BS002 only one watchdogregister for CDIAS and DIAS (IM)
        END_IF;
      END_IF;

    #IFNDEF MaxWatchdog	// #BS016
    END_IF;
	#ENDIF
  END_IF; //ws005

END_FUNCTION // DiasMasterMain::WdCDIAS
FUNCTION VIRTUAL GLOBAL DiasMasterMain::AddDiasIRQ
  VAR_INPUT
    Place		  : USINT;
    ActionPtr	: pVoid;
    thisptr		: pVoid;
  END_VAR
  VAR_OUTPUT
    ok		    : USINT;
  END_VAR

	ok := 0;
	IF IRQDias.anz <= 7 THEN // only 8 Irqs are possible
		IRQDias.data[IRQDias.anz$SINT].ActionPtr	:= ActionPtr;// #BS016
		IRQDias.data[IRQDias.anz$SINT].ThisPtr	:= thisptr;// #BS016
		IF OS_DiasIRQ(TO_USINT(place), #DiasIRQCall() , #IRQDias.data[IRQDias.anz$SINT]) = 0 THEN// #BS016
			ok := 1;
			IRQDias.anz += 1;
		END_IF;
		IF DiasType = 2 THEN
			// #BS001
#ifdef HWC_LogError
      HWC_LogError(thisptr$pVirtualBase, "@0007 (DiasMasterMain::AddDiasIRQ) Interupts on DiasBus with intelligent master are not supported !!! Configurationerror in this object");
#else
			Trace("Interupts on DiasBus with intelligent master are not supported !!! Configurationerror in object:");
#endif
			ok := 0; // only till os gives right value back
		END_IF;
	ELSE // #BS010
#ifdef HWC_LogError
      HWC_LogError(thisptr$pVirtualBase, "@0008 (DiasMasterMain::AddDiasIRQ) Diasinterruptlist is full !! No IRQ for this object");
#else
		Trace("Diasinterruptlist is full !! No IRQ for object:"); // #BS010
#endif
	END_IF;

END_FUNCTION
//[#DEUTSCH]
//[>irqnr]0..IRQ I/O (IRQ PIN C3) | 1..IRQ Comunication (GP2 PIN A10)
FUNCTION VIRTUAL GLOBAL DiasMasterMain::AddCDiasIRQ
  VAR_INPUT
    irqnr		: USINT;
    ActionPtr	: pVoid;
    thisp		: pVoid;
  END_VAR
  VAR_OUTPUT
    ok		: USINT;
  END_VAR

	ok := 0;
	IF CDiasIRQpossible THEN // if possible
		IF OS_INSTALL_CDIAS_IRQ(irqnr, ActionPtr, thisp) = 0 THEN
			ok := 1;
		END_IF;
	END_IF;

END_FUNCTION

#ifdef _LSL_TARGETARCH_X86
FUNCTION AWL DiasMasterMain::DiasIRQCall
	VAR_INPUT
    Station		: UINT;
    ThisIn		: ^USINT;
	END_VAR

//hier die Bedeutung des Registers EBP in Bezug auf den Stack:
//
//+-----------+
//|   param1  |
//+-----------+
//|   param0  | <--- this is [ebp + 8] ( assuming mov ebp, esp )
//+-----------+
//|ret_address|
//+-----------+
//|    ebp    |
//+-----------+ <--- esp
//
//Also, auf EBP + 8 beginnt der 1. Übergabeparameter. In deinem Fall die
//Stationsnummer. Diese wird nur mit 16 Bit Länge auf den Stack gepusht. D.h.,
//der nächste Übergabeparameter beginnt auf EBP + 10. Hier handelt es sich
//dann um ThisIn.
//
//Auf einer 32-Bit-Maschine sollten Übergabeparameter eigentlich immer mit
//32-Bit auf dem Stack landen, da es ansonsten zu einem Misaligned
//Stack-Pointer kommen kann.

// to get a standard interface

	L.EDI		(EBP+10)
	L.ESI		(EDI+oneIRQ.ThisPtr)
	CALL		(EDI+oneIRQ.ActionPtr)

END_FUNCTION
#else
#pragma warning(disable:73 )
FUNCTION DiasMasterMain::DiasIRQCall
	VAR_INPUT
		Station 	: UINT;
		ThisIn 	  : ^USINT;
	END_VAR
  #pragma warning(Default:73)

#ifdef DM_DEBUG_ARM
  // This method is not supported with ARM
  ((0)$^USINT)^ := 0;
#endif

  //LanSte Method is not needed for ARM CPU

END_FUNCTION
#endif

#ifdef _LSL_TARGETARCH_ARM
FUNCTION VIRTUAL GLOBAL DiasMasterMain::RtWorkIMCIPC
  VAR_INPUT
    EAX		: UDINT;
  END_VAR
  VAR_OUTPUT
    state		: UDINT;
  END_VAR
  VAR
    Temp      : DINT;
    pHandle   : ^OneHandle;
    i     :    UDINT;
  //-------------------------------------Profiler Start----------------------------------------------
  #ifdef DiasMasterC_Profiler
    MuSecTime : UDINT;
  END_VAR

  MuSecTime := OS_ReadMicroSec();
  //Anfangsdelay abwarten
	if MuSecTime - DMC_Time_RT.init > DM_ProfilerDelay then
    DMC_Time_RT.start  := MuSecTime;    //Startzeit nehmen
    DMC_Time_RT.initfl := FALSE;        //Initflag löschen
  else
    DMC_Time_RT.initfl := TRUE;         //Initflag setzen
  end_if;
//-------------------------------------Profiler End------------------------------------------------
#else
  END_VAR
#endif

  if (ImOff = FALSE) then
    if (b_TaskTimeCorrected = 0) | (CDIASSync + 3)^ then
      if HwControl = 0 then
        SendSync();
      end_if;

      //look if Rt program of IM is finished
      if (ops.SysState = C_RUNRAM) & (_IOSegment$^USINT + DmUserData + 3)^ then
        ud_ErrorCountTimeSliceEnd += 1;
        if us_FirstTimeSliceEnd = 0 then
          us_FirstTimeSliceEnd := 1;
        end_if;
      end_if;

      //Reset Byte to find out if Rt of IM starts while Rt of DM is running
      (_IOSegment$^USINT + DmUserData + 4)^ := 0;

      case RtSSW of

          // ***********************************************************
          //   we have to wait that the PLL is locked before we start
          // ***********************************************************
        0:

          if Release <> 16#FFFFFFFF then
            if ((_IOSegment$^USINT + DmPllSyncState)^ AND DmPLLisLock) = DmPLLisLock then
              StartRealtimeProg();
              RtSSW += 1;
              LogRtSSW();
            end_if;

            // Start it always to keep the moduls alive
            (_IOSegment$^USINT + DmState)^ := (_IOSegment$^USINT + DmState)^ OR 16#10;
          end_if;

          // **********************************************************
          //  now we are starting the RTProg
          // **********************************************************
        1:

          StartRealtimeProg();
          RtSSW += 1;
          LogRtSSW();

          // ****************************************************************
          //  now we have to move the startpoint till we are 50usec before
          // ****************************************************************
        2:

          if us_MuSecMode then
            Temp := RtInterval - (ud_DelayRealtime / (DmTmrResso * 1000))$DINT - DmTimeReserveIM;
          else
            Temp := RtInterval - (ud_DelayRealtime / (DmTmrResso * 1000))$DINT - (DmTimeReserveIM + 1);
          end_if;

          (_IOSegment$^USINT + DmPllSyncDel)^ := Temp$USINT;
          ui_RtStartPoint := Temp$UINT * DmTmrResso;
          RtSSW += 1;
          LogRtSSW();

          // ***********************************************************
          //   read the calculated time
          // ***********************************************************
        3:

          TimeBeforeNextSync := to_uint((_IOSegment$^USINT + DmUserData)^);
          RtSSW += 1;
          LogRtSSW();

          // ***************************************************************
          //   do the refresh of I/O
          // ***************************************************************
        4:

          // get rtload of im
          TimeAtRtPreEnd := to_dint((_IOSegment$^USINT + DmUserData)^) * DmTmrResso;
          Rt_Load := ((TimeAtRtPreEnd - ui_RtStartPoint) * 1000) / sd_PllTimeGlob_us;

          RealtimeReady := TRUE;

          // now take data and call update methods with thispointer
          if HandleNrRT then
            pHandle := #HandlesRT[0];
            for i := 0 to HandleNrRT-1 do
              if pHandle^.Typ AND DmCallProg then
                pHandle^.thisp^.UpdateRt(pHandle^.Address);
              end_if;

              pHandle += sizeof(OneHandle);
            end_for;
          end_if;

          if HwControl = 0 then
            UpdateRtPostScan_IM();
          end_if;

      end_case;

      if (StateCDiasSync AND 1) = 0 then
        StateCDiasSync := (CDIASSync + 2)^;
      end_if;

      WdCDIAS();
    end_if;
  end_if;

  state := READY;

//-------------------------------------Profiler Start----------------------------------------------
#ifdef DiasMasterC_Profiler
  //schaun ob Delayzeit schon abgelaufen ist
  if DMC_Time_RT.initfl = FALSE then
    MuSecTime := OS_ReadMicroSec();

    DMC_Time_RT.stop := MuSecTime;        //Stopzeit speichern

    MuSecTime -= DMC_Time_RT.start;       //Differenz berechnen
    MuSecTime -= DM_CPUconstant;          //Zeit für OS_REadMicroSec - Funktion subtrahieren

    DMC_Time_RT.diff := MuSecTime;        //korr. Differenz speichern
    DMC_Time_RT.sum  += MuSecTime;        //Zur Summe addieren

    DMC_Time_RT.run  += 1;                //Durchlaufzähler erhöhen

    if MuSecTime < DMC_Time_RT._min then
      DMC_Time_RT._min := MuSecTime;      //Minimalzeit speichern
    end_if;

    if MuSecTime > DMC_Time_RT._max then
      DMC_Time_RT._max := MuSecTime;      //Maximalzeit speichern
    end_if;

    //Durchschnitt berechnen
    //*100 damit wir 2 Kommastellen haben
    DMC_Time_RT.avg := DMC_Time_RT.sum * 100 / DMC_Time_RT.run;
  end_if;

#endif
//-------------------------------------Profiler End------------------------------------------------
END_FUNCTION

#else

FUNCTION AWL VIRTUAL GLOBAL DiasMasterMain::RtWorkIMCIPC
  VAR_INPUT
    EAX		: UDINT;
  END_VAR
  VAR_OUTPUT
    state		: UDINT;
  END_VAR

//#wp001
//============================ Profiler start======================================================
#ifdef  DiasMasterC_Profiler
	CLI											//damit keine Interrupts die Messung stören
	push 		  edi
	push 		  eax
	l.edi 		_LSL_POS
	l.edi 		( edi + DM_LSLPOS_SYSTIME )
	l.edi 		( edi + DM_LSLSYSTIME_MICROSEC )
	call		  edi								//OS_ReadMicroSec - Funktion aufrufen
	l.ebx		  eax
	sub.ebx		DMC_Time_RT.init					//Anfangsdelay abwarten
	cmp.ebx		DM_ProfilerDelay
	jle			  LABEL_DMCPREEND
	s.eax 		DMC_Time_RT.start					//Startzeit nehmen
	x.cl		  cl
	s.cl		  DMC_Time_RT.initfl				//Initflag löschen
	jmp 		  LABEL_DMCstartfunc

LABEL_DMCPREEND
	l.b		    DMC_Time_RT.initfl,1					//Initflag setzen

LABEL_DMCstartfunc
	pop 		  eax
	pop 		  edi
#endif
//============================ Profiler end========================================================

	CMP.B			ImOff,1
	JE				RT_End1

  cmp.b     b_TaskTimeCorrected, 1
  jne       LABEL_AfterTaskCheck

  // task selector over fpga bit => to ensure synchronity
  l.edi     CDIASSync
  l         (edi + 3)
  cmp.al    0
  jz        RT_End1

LABEL_AfterTaskCheck

	//#SR014 start
	cmp.d			HwControl, 1
	je				LABEL_EndPllSync

	call			SendSync
	//#SR014 end

LABEL_EndPllSync	//#SR013

	//#SR010 start
	cmp.w			ops.SysState,1					//look if CPU is in RunRam
	jne				LABEL_Continue

 	l.edi			_IOSegment						//#SR014
	l.bl			( edi + DmUserData + 3 )		//look if Rt program of IM is finished
	o.bl			bl
	jz				LABEL_Continue
	inc.d			ud_ErrorCountTimeSliceEnd
	cmp.b			us_FirstTimeSliceEnd,0
	jne				LABEL_Continue

	l.b				us_FirstTimeSliceEnd,1
LABEL_Continue
  l.edi			_IOSegment						//#SR014
	l.b				( edi + DmUserData + 4 ), 0		//Reset Byte to find out if Rt of IM starts while Rt of DM is running
	//#SR010 end

	lzxb.eax	RtSSW		//ws005
	shl.eax		3             //ws005: save some time here
	add.eax		#RtSel
	jmp			  eax

RtSel
	jmp			WaitForSync			// 0 : wait till PLL in locked
	rcl.eax 	0					//ws005: simple placeholder (does really nothing)
	jmp			weAreSync			// 1 : wait one period to get a right time
	rcl.eax 	0					//ws005: simple placeholder (does really nothing)
	jmp			MovStartPoint		// 2 : mov start point to the right pos
	rcl.eax 	0					//ws005: simple placeholder (does really nothing)
	jmp			readpoint           // 3 : read one time the point
	rcl.eax 	0					//ws005: simple placeholder (does really nothing)
	jmp			RtRefresh			// 4 : do the realtime refresh

// ***************************************************************
//   do the refresh of I/O
// ***************************************************************

RtRefresh

// *************************************************
//  read the time point
// *************************************************
	lzxb.eax	(edi+DmUserData)
	imul.ax		ax,DmTmrResso
	s.eax 		TimeAtRtPreEnd

	//#SR009
	//***********calculate Rt - usage rate***********************
	lzxw.ebx	ui_RtStartPoint
	sub.eax		ebx
	imul.eax	eax,1000
	x.edx		  edx
	l.ebx		  sd_PllTimeGlob_us
	div			  ebx
	s.eax		  Rt_Load
	//#SR009

// **************************************************
//  now take data and call update function with thisp
// **************************************************
	l.b			  RealtimeReady,1		//ws005

	l.ebx		  #HandlesRt
	lzxw.ecx	HandleNrRt
	jecxz		  LABEL_RtPostScan		//#SR010 RT_end    //NoRtProg  //ws005

HandleLoopRt
	test.w		(ebx+OneHandle.Typ),DmCallProg
	jz			  NextHandleRt
